	    // Condition to request disable send
	    #s_Ext_Req_Disable_Send := #i_External_Request.Request_Disable_Send;

	    // Condition to request disable receive
	    #s_Ext_Req_Disable_Recv := #i_External_Request.Request_Disable_Receive OR #i_Command.Man_Mode;

	    // Condition to request reset engergy saving
	    #s_Ext_Req_Rest_ESave := #i_External_Request.Request_Reset_EnergySave OR #io_Global.Common_Setting.Disable_Energy_Saving OR #i_Command.Cmd_Reset_ESave OR #s_FB_EQP_PEC_Position.s_PEC_Filter;

	    // Condition to request clear flow interface data
	    #s_Ext_Req_Clear_Data := #i_External_Request.Request_Clear_Data OR (#i_Command.Man_Clear AND #i_Command.Man_Mode);
	END_REGION

	REGION NETWORK DA: Equipment Layer - Basic
	    #s_FB_EQP_Transport(i_Enable                 := #io_System_Control.Enable,
	                        i_IO_Available           := #io_System_Control.IO_Available,
	                        i_Safety_OK              := #io_System_Control.Safety_OK,
	                        i_CMD_Reset              := #io_System_Control.OS_Reset,
	                        i_CMD_Start              := #io_System_Control.OS_Start,
	                        i_CMD_Controlled_Stop    := #io_System_Control.Controlled_Stop,
	                        i_End_PEC_Latch          := #s_PE_Position_Latch,
	                        i_Manual_Run             := #i_Command.Man_Run AND #i_Command.Man_Mode,
	                        i_CFG_Slave_Conveyor     := #i_Setting.Base_Conveyor.Slave_Mode,
	                        i_CFG_Enable_DieForward  := #i_Setting.Base_Conveyor.Enable_DieForward,
	                        i_Delay_Waiting_Item     := #i_Setting.Base_Conveyor.Delay_Waiting_Item,
	                        i_Delay_Dieback          := #i_Setting.Base_Conveyor.Delay_Dieback,
	                        i_Delay_Startup          := #i_Setting.Base_Conveyor.Delay_Startup,
	                        i_Delay_Finish_Handover  := #i_Setting.Base_Conveyor.Delay_Finish_Handover,
	                        i_Delay_Energysave       := #i_Setting.Base_Conveyor.Delay_Energysave,
	                        i_Delay_Cascade_Startup  := #i_Setting.Base_Conveyor.Delay_Cascade_Startup,
	                        i_Delay_Cascade_Shutdown := #i_Setting.Base_Conveyor.Delay_Cascade_Shutdown,
	                        i_Delay_Motor_Startup    := 0,
	                        i_Minimum_Gap            := #i_Setting.Flow_Control.Minimum_Gap,
	                        i_Minimum_Head_To_Head   := #i_Setting.Flow_Control.Minimum_Head_To_Head,
	                        i_Ext_Req_Stop           := #s_Ext_Req_Stop,
	                        i_Ext_Req_Halt           := #s_Ext_Req_Halt,
	                        i_Ext_Req_Dis_Send       := #s_Ext_Req_Disable_Send,
	                        i_Ext_Req_Dis_Recv       := #s_Ext_Req_Disable_Recv,
	                        i_Ext_Req_Rst_ESave      := #s_Ext_Req_Rest_ESave,
	                        i_Ext_Req_Clear_Data     := #s_Ext_Req_Clear_Data,
	                        o_Ready_To_Start         => #io_System_Control.Ready_To_Start,
	                        o_ST_Safety_Stop         => #o_General_Status.Safety_Stop,
	                        o_ST_Items               => #o_General_Status.Items,
	                        o_ST_Die_Back            => #o_General_Status.Die_Back,
	                        o_ST_Motor_Running       => #o_General_Status.Motor_Running,
	                        o_ST_Started             => #o_General_Status.Started,
	                        o_ST_Energy_Saving       => #o_General_Status.Energy_Saving,
	                        o_MTR_Run                => #s_CMD_Motor,
	                        io_Global                := #io_Global,
	                        io_FIF_Upstream          := #io_FIF_Upstream,
	                        io_FIF                   := #io_FIF,
	                        io_FIF_Downstream        := #io_FIF_Downstream);
	END_REGION

	REGION NETWORK EA: Hardware Layer - Interroll MultiControl 1
	    #s_Speed_Select := #i_External_Request.Request_Speed;

	    #s_FB_HW_MultiControl_U01(i_IO_Available            := #io_System_Control.IO_Available,
	                              i_Safety_OK               := #io_System_Control.Safety_OK,
	                              i_CMD_Reset               := #io_System_Control.OS_Reset,
	                              i_CMD_Clear_Stat          := #io_System_Control.OS_Clear_Statistics,
	                              i_HW_Setting              := #i_Setting.Hardware_U01,
	                              i_CFG_Motor_Switch_Time   := 500,
	                              i_CMD_Select_Speed        := #s_Speed_Select,
	                              i_CMD_Motor_Run           := #s_CMD_Motor,
	                              i_CMD_Motor_Reverse       := #s_CMD_Motor_Reverse,
	                              o_Ready_To_Reset          => #t_HW_VFD_U01_Ready_To_Reset,
	                              o_Req_Halt                => #s_HW_U01_Req_Halt,
	                              o_ER_Motor_1_Fault        => #t_ER_Motor_U01_Fault,
	                              o_ER_Motor_2_Fault        => #t_ER_Motor_U02_Fault,
	                              o_ER_Motor_3_Fault        => #t_ER_Motor_U03_Fault,
	                              o_ER_Motor_4_Fault        => #t_ER_Motor_U04_Fault,
	                              o_Speed_Selected          => #io_FIF.Speed,
	                              o_Diagnostics             => #o_Diagnostics.Hardware_U01,
	                              io_Global                 := #io_Global,
	                              io_MultiControl_Interface := #io_MultiControl_U01_IO);

	    IF #i_Setting.Hardware_U01.RD1_Motor_Number > 0 AND #i_Setting.Hardware_U01.RD1_Motor_Number <= 16 THEN
	        #t_ER_Motor_Fault[#i_Setting.Hardware_U01.RD1_Motor_Number] := #t_ER_Motor_U01_Fault;
	    END_IF;

	    IF #i_Setting.Hardware_U01.RD2_Motor_Number > 0 AND #i_Setting.Hardware_U01.RD2_Motor_Number <= 16 THEN
	        #t_ER_Motor_Fault[#i_Setting.Hardware_U01.RD2_Motor_Number] := #t_ER_Motor_U02_Fault;
	    END_IF;

	    IF #i_Setting.Hardware_U01.RD3_Motor_Number > 0 AND #i_Setting.Hardware_U01.RD3_Motor_Number <= 16 THEN
	        #t_ER_Motor_Fault[#i_Setting.Hardware_U01.RD3_Motor_Number] := #t_ER_Motor_U03_Fault;
	    END_IF;

	    IF #i_Setting.Hardware_U01.RD4_Motor_Number > 0 AND #i_Setting.Hardware_U01.RD4_Motor_Number <= 16 THEN
	        #t_ER_Motor_Fault[#i_Setting.Hardware_U01.RD4_Motor_Number] := #t_ER_Motor_U04_Fault;
	    END_IF;
	END_REGION

	REGION NETWORK EB: Hardware Layer - Interroll MultiControl 2
	    #s_Speed_Select := #i_External_Request.Request_Speed;

	    #s_FB_HW_MultiControl_U02(i_IO_Available            := #io_System_Control.IO_Available,
	                              i_Safety_OK               := #io_System_Control.Safety_OK,
	                              i_CMD_Reset               := #io_System_Control.OS_Reset,
	                              i_CMD_Clear_Stat          := #io_System_Control.OS_Clear_Statistics,
	                              i_HW_Setting              := #i_Setting.Hardware_U02,
	                              i_CFG_Motor_Switch_Time   := 500,
	                              i_CMD_Select_Speed        := #s_Speed_Select,
	                              i_CMD_Motor_Run           := #s_CMD_Motor,
	                              i_CMD_Motor_Reverse       := #s_CMD_Motor_Reverse,
	                              o_Ready_To_Reset          => #t_HW_VFD_U02_Ready_To_Reset,
	                              o_Req_Halt                => #s_HW_U02_Req_Halt,
	                              o_ER_Motor_1_Fault        => #t_ER_Motor_U01_Fault,
	                              o_ER_Motor_2_Fault        => #t_ER_Motor_U02_Fault,
	                              o_ER_Motor_3_Fault        => #t_ER_Motor_U03_Fault,
	                              o_ER_Motor_4_Fault        => #t_ER_Motor_U04_Fault,
	                              o_Diagnostics             => #o_Diagnostics.Hardware_U02,
	                              io_Global                 := #io_Global,
	                              io_MultiControl_Interface := #io_MultiControl_U02_IO);

	    IF #i_Setting.Hardware_U02.RD1_Motor_Number > 0 AND #i_Setting.Hardware_U02.RD1_Motor_Number <= 16 THEN
	        #t_ER_Motor_Fault[#i_Setting.Hardware_U02.RD1_Motor_Number] := #t_ER_Motor_U01_Fault;
	    END_IF;

	    IF #i_Setting.Hardware_U02.RD2_Motor_Number > 0 AND #i_Setting.Hardware_U02.RD2_Motor_Number <= 16 THEN
	        #t_ER_Motor_Fault[#i_Setting.Hardware_U02.RD2_Motor_Number] := #t_ER_Motor_U02_Fault;
	    END_IF;

	    IF #i_Setting.Hardware_U02.RD3_Motor_Number > 0 AND #i_Setting.Hardware_U02.RD3_Motor_Number <= 16 THEN
	        #t_ER_Motor_Fault[#i_Setting.Hardware_U02.RD3_Motor_Number] := #t_ER_Motor_U03_Fault;
	    END_IF;

	    IF #i_Setting.Hardware_U02.RD4_Motor_Number > 0 AND #i_Setting.Hardware_U02.RD4_Motor_Number <= 16 THEN
	        #t_ER_Motor_Fault[#i_Setting.Hardware_U02.RD4_Motor_Number] := #t_ER_Motor_U04_Fault;
	    END_IF;
	END_REGION

	REGION NETWORK EA: Hardware Layer - Interroll MultiControl 3
	    #s_Speed_Select := #i_External_Request.Request_Speed;

	    #s_FB_HW_MultiControl_U03(i_IO_Available            := #io_System_Control.IO_Available,
	                              i_Safety_OK               := #io_System_Control.Safety_OK,
	                              i_CMD_Reset               := #io_System_Control.OS_Reset,
	                              i_CMD_Clear_Stat          := #io_System_Control.OS_Clear_Statistics,
	                              i_HW_Setting              := #i_Setting.Hardware_U03,
	                              i_CFG_Motor_Switch_Time   := 500,
	                              i_CMD_Select_Speed        := #s_Speed_Select,
	                              i_CMD_Motor_Run           := #s_CMD_Motor,
	                              i_CMD_Motor_Reverse       := #s_CMD_Motor_Reverse,
	                              o_Ready_To_Reset          => #t_HW_VFD_U03_Ready_To_Reset,
	                              o_Req_Halt                => #s_HW_U03_Req_Halt,
	                              o_ER_Motor_1_Fault        => #t_ER_Motor_U01_Fault,
	                              o_ER_Motor_2_Fault        => #t_ER_Motor_U02_Fault,
	                              o_ER_Motor_3_Fault        => #t_ER_Motor_U03_Fault,
	                              o_ER_Motor_4_Fault        => #t_ER_Motor_U04_Fault,
	                              o_Diagnostics             => #o_Diagnostics.Hardware_U03,
	                              io_Global                 := #io_Global,
	                              io_MultiControl_Interface := #io_MultiControl_U03_IO);

	    IF #i_Setting.Hardware_U03.RD1_Motor_Number > 0 AND #i_Setting.Hardware_U03.RD1_Motor_Number <= 16 THEN
	        #t_ER_Motor_Fault[#i_Setting.Hardware_U03.RD1_Motor_Number] := #t_ER_Motor_U01_Fault;
	    END_IF;

	    IF #i_Setting.Hardware_U03.RD2_Motor_Number > 0 AND #i_Setting.Hardware_U03.RD2_Motor_Number <= 16 THEN
	        #t_ER_Motor_Fault[#i_Setting.Hardware_U03.RD2_Motor_Number] := #t_ER_Motor_U02_Fault;
	    END_IF;

	    IF #i_Setting.Hardware_U03.RD3_Motor_Number > 0 AND #i_Setting.Hardware_U03.RD3_Motor_Number <= 16 THEN
	        #t_ER_Motor_Fault[#i_Setting.Hardware_U03.RD3_Motor_Number] := #t_ER_Motor_U03_Fault;
	    END_IF;

	    IF #i_Setting.Hardware_U03.RD4_Motor_Number > 0 AND #i_Setting.Hardware_U03.RD4_Motor_Number <= 16 THEN
	        #t_ER_Motor_Fault[#i_Setting.Hardware_U03.RD4_Motor_Number] := #t_ER_Motor_U04_Fault;
	    END_IF;
	END_REGION

	REGION NETWORK EA: Hardware Layer - Interroll MultiControl 4
	    #s_Speed_Select := #i_External_Request.Request_Speed;

	    #s_FB_HW_MultiControl_U04(i_IO_Available            := #io_System_Control.IO_Available,
	                              i_Safety_OK               := #io_System_Control.Safety_OK,
	                              i_CMD_Reset               := #io_System_Control.OS_Reset,
	                              i_CMD_Clear_Stat          := #io_System_Control.OS_Clear_Statistics,
	                              i_HW_Setting              := #i_Setting.Hardware_U04,
	                              i_CFG_Motor_Switch_Time   := 500,
	                              i_CMD_Select_Speed        := #s_Speed_Select,
	                              i_CMD_Motor_Run           := #s_CMD_Motor,
	                              i_CMD_Motor_Reverse       := #s_CMD_Motor_Reverse,
	                              o_Ready_To_Reset          => #t_HW_VFD_U04_Ready_To_Reset,
	                              o_Req_Halt                => #s_HW_U04_Req_Halt,
	                              o_ER_Motor_1_Fault        => #t_ER_Motor_U01_Fault,
	                              o_ER_Motor_2_Fault        => #t_ER_Motor_U02_Fault,
	                              o_ER_Motor_3_Fault        => #t_ER_Motor_U03_Fault,
	                              o_ER_Motor_4_Fault        => #t_ER_Motor_U04_Fault,
	                              o_Diagnostics             => #o_Diagnostics.Hardware_U04,
	                              io_Global                 := #io_Global,
	                              io_MultiControl_Interface := #io_MultiControl_U04_IO);

	    IF #i_Setting.Hardware_U04.RD1_Motor_Number > 0 AND #i_Setting.Hardware_U04.RD1_Motor_Number <= 16 THEN
	        #t_ER_Motor_Fault[#i_Setting.Hardware_U04.RD1_Motor_Number] := #t_ER_Motor_U01_Fault;
	    END_IF;

	    IF #i_Setting.Hardware_U04.RD2_Motor_Number > 0 AND #i_Setting.Hardware_U04.RD2_Motor_Number <= 16 THEN
	        #t_ER_Motor_Fault[#i_Setting.Hardware_U04.RD2_Motor_Number] := #t_ER_Motor_U02_Fault;
	    END_IF;

	    IF #i_Setting.Hardware_U04.RD3_Motor_Number > 0 AND #i_Setting.Hardware_U04.RD3_Motor_Number <= 16 THEN
	        #t_ER_Motor_Fault[#i_Setting.Hardware_U04.RD3_Motor_Number] := #t_ER_Motor_U03_Fault;
	    END_IF;

	    IF #i_Setting.Hardware_U04.RD4_Motor_Number > 0 AND #i_Setting.Hardware_U04.RD4_Motor_Number <= 16 THEN
	        #t_ER_Motor_Fault[#i_Setting.Hardware_U04.RD4_Motor_Number] := #t_ER_Motor_U04_Fault;
	    END_IF;
	END_REGION

	REGION NETWORK: Copy Motor Alarm to Status

	    #o_Status.ER_Motor_1_Fault := #t_ER_Motor_Fault[1];
	    #o_Status.ER_Motor_2_Fault := #t_ER_Motor_Fault[2];
	    #o_Status.ER_Motor_3_Fault := #t_ER_Motor_Fault[3];
	    #o_Status.ER_Motor_4_Fault := #t_ER_Motor_Fault[4];
	    #o_Status.ER_Motor_5_Fault := #t_ER_Motor_Fault[5];
	    #o_Status.ER_Motor_6_Fault := #t_ER_Motor_Fault[6];
	    #o_Status.ER_Motor_7_Fault := #t_ER_Motor_Fault[7];
	    #o_Status.ER_Motor_8_Fault := #t_ER_Motor_Fault[8];
	    #o_Status.ER_Motor_9_Fault := #t_ER_Motor_Fault[9];
	    #o_Status.ER_Motor_10_Fault := #t_ER_Motor_Fault[10];
	    #o_Status.ER_Motor_11_Fault := #t_ER_Motor_Fault[11];
	    #o_Status.ER_Motor_12_Fault := #t_ER_Motor_Fault[12];
	    #o_Status.ER_Motor_13_Fault := #t_ER_Motor_Fault[13];
	    #o_Status.ER_Motor_14_Fault := #t_ER_Motor_Fault[14];
	    #o_Status.ER_Motor_15_Fault := #t_ER_Motor_Fault[15];
	    #o_Status.ER_Motor_16_Fault := #t_ER_Motor_Fault[16];

	END_REGION

	REGION NETWORK: Diagnositcs
	    #o_Diagnostics.RTS := #io_FIF.RTS;
	    #o_Diagnostics.TIP := #io_FIF.TIP;
	    #o_Diagnostics.Downstream_RTR := #io_FIF_Downstream.RTR;
	    #o_Diagnostics.Displacement := #io_FIF.Displacement;
	    #o_Diagnostics.Items_Count := MAX_UDINT(IN1 := #t_PEC_Position_Items, IN2 := #t_PEC_Trigger_Items);
	END_REGION

	REGION NETWORK FA: Make Generate Status
	    #o_Status.OL_Maintenance_Mode := #i_Command.Man_Mode;

	    #o_General_Status.Safety_Stop := NOT #io_System_Control.Safety_OK;
	    #o_General_Status.Off_Line := #o_Status.OL_Maintenance_Mode;
	    #o_General_Status.Manual := FALSE;
	    #o_General_Status.Error := #o_Status.ER_Motor_1_Fault
	    OR #o_Status.ER_Motor_2_Fault
	    OR #o_Status.ER_Motor_3_Fault
	    OR #o_Status.ER_Motor_4_Fault
	    OR #o_Status.ER_Motor_5_Fault
	    OR #o_Status.ER_Motor_6_Fault
	    OR #o_Status.ER_Motor_7_Fault
	    OR #o_Status.ER_Motor_8_Fault
	    OR #o_Status.ER_Motor_9_Fault
	    OR #o_Status.ER_Motor_10_Fault
	    OR #o_Status.ER_Motor_11_Fault
	    OR #o_Status.ER_Motor_12_Fault
	    OR #o_Status.ER_Motor_13_Fault
	    OR #o_Status.ER_Motor_14_Fault
	    OR #o_Status.ER_Motor_15_Fault
	    OR #o_Status.ER_Motor_16_Fault;
	    #o_General_Status.Jam := #o_Status.ER_PE1_Blockage OR #o_Status.ER_PE2_Blockage;
	END_REGION

	REGION NETWORK EA: System Feedback State
	    #io_System_Control.Ready_To_Reset := #t_PEC_Position_Ready_To_Reset
	    OR #t_PEC_Trigger_Ready_To_Reset
	    OR #t_HW_VFD_U01_Ready_To_Reset
	    OR #t_HW_VFD_U02_Ready_To_Reset
	    OR #t_HW_VFD_U03_Ready_To_Reset
	    OR #t_HW_VFD_U04_Ready_To_Reset;
	END_REGION
END_FUNCTION_BLOCK

TYPE "UDT_GL2S_IO"
VERSION : 0.1
   STRUCT
      IsCleared : Bool;
   END_STRUCT;

END_TYPE

TYPE "UDT_Conv_Triple_G115D_Status"
VERSION : 0.1
   STRUCT
      OL_Maintenance_Mode : Bool;   // Maintenance mode on
      ER_PE1_Blockage : Bool;   // PE1 blockage
      ER_PE2_Blockage : Bool;   // PE2 blockage
      ER_U01_VFD_PN_NotPresent : Bool;   // VFD 1# not present on profinet network
      ER_U01_VFD_PN_Error : Bool;   // VFD 1# has error profinet network
      ER_U01_VFD_Fault : Bool;   // VFD 1# has error
      WN_U01_VFD_Alarm : Bool;   // VFD 1# has an warning
      ER_U01_VFD_STO_Active : Bool;   // VFD 1# STO is active
      WN_U01_No_MemoryCard : Bool;   // Memory card is missing
      ER_U02_VFD_PN_NotPresent : Bool;   // VFD 2# not present on profinet network
      ER_U02_VFD_PN_Error : Bool;   // VFD 2# has error profinet network
      ER_U02_VFD_Fault : Bool;   // VFD 2# has error
      WN_U02_VFD_Alarm : Bool;   // VFD 2# has an warning
      ER_U02_VFD_STO_Active : Bool;   // VFD 2# STO is active
      WN_U02_No_MemoryCard : Bool;   // Memory card is missing
      ER_U03_VFD_PN_NotPresent : Bool;   // VFD 3# not present on profinet network
      ER_U03_VFD_PN_Error : Bool;   // VFD 3# has error profinet network
      ER_U03_VFD_Fault : Bool;   // VFD 3# has error
      WN_U03_VFD_Alarm : Bool;   // VFD 3# has an warning
      ER_U03_VFD_STO_Active : Bool;   // VFD 3# STO is active
      WN_U03_No_MemoryCard : Bool;   // Memory card is missing
      Spare_2_5 : Bool;   // Spare_2_5
      Spare_2_6 : Bool;   // Spare_2_6
      Spare_2_7 : Bool;   // Spare_2_7
      Spare_3_0 : Bool;   // Spare_3_0
      Spare_3_1 : Bool;   // Spare_3_1
      Spare_3_2 : Bool;   // Spare_3_2
      Spare_3_3 : Bool;   // Spare_3_3
      Spare_3_4 : Bool;   // Spare_3_4
      Spare_3_5 : Bool;   // Spare_3_5
      Spare_3_6 : Bool;   // Spare_3_6
      Spare_3_7 : Bool;   // Spare_3_7
      U01_FaultCode : Word;   // VFD 1# fault code
      U01_AlarmCode : Word;   // VFD 1# alarm code
      U02_FaultCode : Word;   // VFD 2# fault code
      U02_AlarmCode : Word;   // VFD 2# alarm code
      U03_FaultCode : Word;   // VFD 3# fault code
      U03_AlarmCode : Word;   // VFD 3# alarm code
   END_STRUCT;

END_TYPE

FUNCTION_BLOCK "FB_Conv_SWS"
{ S7_Optimized_Access := 'TRUE' }
VERSION : 0.1
   VAR_INPUT
      i_New_Item_Present : Bool;
      i_CMD_Divert_Left : Bool;
      i_CMD_Divert_Straight : Bool;
      i_CMD_Divert_Right : Bool;
      i_Setting : "UDT_Conv_SWS_Setting";
      i_External_Request : "UDT_External_Request";
      i_U401_Additional_HW_ID : HW_SUBMODULE;
      i_U401_Telegram_HW_ID : HW_SUBMODULE;
      i_U411_Additional_HW_ID : HW_SUBMODULE;
      i_U411_Telegram_HW_ID : HW_SUBMODULE;
      i_U421_Additional_HW_ID : HW_SUBMODULE;
      i_U421_Telegram_HW_ID : HW_SUBMODULE;
      i_U431_Additional_HW_ID : HW_SUBMODULE;
      i_U431_Telegram_HW_ID : HW_SUBMODULE;
      i_U441_Additional_HW_ID : HW_SUBMODULE;
      i_U441_Telegram_HW_ID : HW_SUBMODULE;
      i_U451_Additional_HW_ID : HW_SUBMODULE;
      i_U451_Telegram_HW_ID : HW_SUBMODULE;
      i_U461_Additional_HW_ID : HW_SUBMODULE;
      i_U461_Telegram_HW_ID : HW_SUBMODULE;
      i_U471_Additional_HW_ID : HW_SUBMODULE;
      i_U471_Telegram_HW_ID : HW_SUBMODULE;
      i_U481_Additional_HW_ID : HW_SUBMODULE;
      i_U481_Telegram_HW_ID : HW_SUBMODULE;
      i_Roller_Gateway_Input_HW_ID : HW_ANY;
      i_Roller_Gateway_Output_HW_ID : HW_ANY;
   END_VAR

   VAR_OUTPUT
      o_Status : "UDT_Conv_SWS_Status";
      o_General_Status : "UDT_General_Status";
   END_VAR

   VAR_IN_OUT
      io_Global : "UDT_Global";
      io_System_Control : "UDT_System_Control";
      io_Interface : "UDT_SWS_Interface";
      io_Gateway_Interface : "UDT_NT100_Interface";
      io_Command : "UDT_Conv_SWS_Command";
      io_FIF_Upstream : "UDT_Flow_Interface";
      io_FIF : "UDT_Flow_Interface";
      io_FIF_Downstream : "UDT_Flow_Interface";
   END_VAR

   VAR
      s_FB_Displacement_AccDec : "FB_Displacement_AccDec";
      s_FB_SWS_Roller_Interface : "FB_HW_SWS_Roller_Interface";
      s_FB_EQP_Transport : "FB_EQP_Transport";
      s_Trigger_FB_EQP_PEC_Position : "FB_EQP_PEC_Position";
      s_FB_SWS_Array_Control : "FB_SWS_Array_Control";
      s_U401_FB_SWS_EQP_Servo { S7_SetPoint := 'False'} : "FB_HW_SWS_S210";
      s_U411_FB_SWS_EQP_Servo { S7_SetPoint := 'False'} : "FB_HW_SWS_S210";
      s_U421_FB_SWS_EQP_Servo { S7_SetPoint := 'False'} : "FB_HW_SWS_S210";
      s_U431_FB_SWS_EQP_Servo { S7_SetPoint := 'False'} : "FB_HW_SWS_S210";
      s_U441_FB_SWS_EQP_Servo { S7_SetPoint := 'False'} : "FB_HW_SWS_S210";
      s_U451_FB_SWS_EQP_Servo { S7_SetPoint := 'False'} : "FB_HW_SWS_S210";
      s_U461_FB_SWS_EQP_Servo { S7_SetPoint := 'False'} : "FB_HW_SWS_S210";
      s_U471_FB_SWS_EQP_Servo { S7_SetPoint := 'False'} : "FB_HW_SWS_S210";
      s_U481_FB_SWS_EQP_Servo { S7_SetPoint := 'False'} : "FB_HW_SWS_S210";
      s_Servo_Array_Command : Array[1..#C_ARRAY_COUNT] of Struct
         CMD_Straight : Bool;
         CMD_Left : Bool;
         CMD_Right : Bool;
      END_STRUCT;
      s_Servo_Status { S7_SetPoint := 'False'} : Array[1..#C_ARRAY_COUNT] of "UDT_SWS_Servo_Status";
      s_Roller_Module_Status { ExternalAccessible := 'False'; ExternalVisible := 'False'; ExternalWritable := 'False'; S7_SetPoint := 'False'} : Array[1..9] of "UDT_SWS_Roller_Module_Status";
      s_Servo_Ready_To_Reset : Array[1..#C_ARRAY_COUNT] of Bool;
   END_VAR
   VAR RETAIN
      s_SW_Actual_Speed { S7_SetPoint := 'True'} : Int;
      s_CMD_Roller_Run : Bool;
      s_Ext_Req_Stop : Bool;
      s_Ext_Req_Halt : Bool;
      s_Ext_Req_Disable_Send : Bool;
      s_Ext_Req_Disable_Recv : Bool;
      s_Ext_Req_Rest_ESave : Bool;
      s_Ext_Req_Clear_Data : Bool;
   END_VAR

   VAR_TEMP
      t_GeoAddr {InstructionName := 'GEOADDR'; LibVersion := '1.0'} : GEOADDR;
      t_Ret_Val_Int : Int;   // Temp: Return Value Int
      t_Delayed_Item_Trigger : Bool;
   END_VAR

   VAR CONSTANT
      C_ARRAY_COUNT : UInt := 9;
   END_VAR


BEGIN
	REGION Conveyor Cycle Displacement
	    #io_FIF.Speed := #i_Setting.Hardware.Roller.Speed_Straight;

	    #s_FB_Displacement_AccDec(i_Conveyor_Speed   := #io_FIF.Speed,
	                              i_Accelaration     := #i_Setting.Hardware.Roller.Acceleration,
	                              i_Decelaration     := #i_Setting.Hardware.Roller.Deceleration,
	                              i_Prev_Cycle_Time  := #io_Global.OB_Prev_Cycle_Time,
	                              i_PPI_Displacement := 0,
	                              i_Section_Run      := #io_FIF.Motor_Run,
	                              o_Motor_On_Speed   => #o_General_Status.Motor_On_Speed,
	                              o_Motor_Stopped    => #io_FIF.Motor_Stopped,
	                              o_Actual_Speed     => #s_SW_Actual_Speed,
	                              o_Displacement     => #io_FIF.Displacement);

	    #o_General_Status.Motor_Stopped := #io_FIF.Motor_Stopped;
	END_REGION

	REGION Roller Hardware Interface
	    #s_FB_SWS_Roller_Interface(i_CFG_HW_Port                := #i_Roller_Gateway_Input_HW_ID,
	                               i_IO_Available               := #io_System_Control.IO_Available,
	                               i_OB_First_Scan              := #io_Global.OS_First_Scan,
	                               i_CMD_Reset                  := #io_System_Control.OS_Reset,
	                               i_CFG_Status_Interval        := #i_Setting.Roller_Interface.Status_Interval,
	                               i_CFG_Num_Of_Comm_Error      := #i_Setting.Roller_Interface.Num_Of_Comm_Error,
	                               i_Sett_Roller_Hardware       := #i_Setting.Hardware.Roller,
	                               i_Roller_Running             := #io_FIF.Motor_Run,
	                               o_ER_Modbus_Initialize_Fault => #o_Status.ER_Modbus_Gateway_Initialize_Fault,
	                               o_ER_Modbus_Com_Error        => #o_Status.ER_Modbus_Gateway_Communication_Fault,
	                               o_Modules_Status             => #s_Roller_Module_Status);

	END_REGION

	REGION Conditions to basic control
	    // Condition to request stop
	    #s_Ext_Req_Stop := #s_Servo_Status[1].ER_PN_NotPresent
	    OR #s_Servo_Status[2].ER_PN_NotPresent
	    OR #s_Servo_Status[3].ER_PN_NotPresent
	    OR #s_Servo_Status[4].ER_PN_NotPresent
	    OR #s_Servo_Status[5].ER_PN_NotPresent
	    OR #s_Servo_Status[6].ER_PN_NotPresent
	    OR #s_Servo_Status[7].ER_PN_NotPresent
	    OR #s_Servo_Status[8].ER_PN_NotPresent
	    OR #s_Servo_Status[9].ER_PN_NotPresent
	    OR #s_Servo_Status[1].ER_Servo_Fault
	    OR #s_Servo_Status[2].ER_Servo_Fault
	    OR #s_Servo_Status[3].ER_Servo_Fault
	    OR #s_Servo_Status[4].ER_Servo_Fault
	    OR #s_Servo_Status[5].ER_Servo_Fault
	    OR #s_Servo_Status[6].ER_Servo_Fault
	    OR #s_Servo_Status[7].ER_Servo_Fault
	    OR #s_Servo_Status[8].ER_Servo_Fault
	    OR #s_Servo_Status[9].ER_Servo_Fault
	    OR #s_Servo_Status[1].ER_Home_Position_Missed
	    OR #s_Servo_Status[2].ER_Home_Position_Missed
	    OR #s_Servo_Status[3].ER_Home_Position_Missed
	    OR #s_Servo_Status[4].ER_Home_Position_Missed
	    OR #s_Servo_Status[5].ER_Home_Position_Missed
	    OR #s_Servo_Status[6].ER_Home_Position_Missed
	    OR #s_Servo_Status[7].ER_Home_Position_Missed
	    OR #s_Servo_Status[8].ER_Home_Position_Missed
	    OR #s_Servo_Status[9].ER_Home_Position_Missed
	    OR #s_Servo_Status[1].ER_STO_Active
	    OR #s_Servo_Status[2].ER_STO_Active
	    OR #s_Servo_Status[3].ER_STO_Active
	    OR #s_Servo_Status[4].ER_STO_Active
	    OR #s_Servo_Status[5].ER_STO_Active
	    OR #s_Servo_Status[6].ER_STO_Active
	    OR #s_Servo_Status[7].ER_STO_Active
	    OR #s_Servo_Status[8].ER_STO_Active
	    OR #s_Servo_Status[9].ER_STO_Active
	    OR #i_External_Request.Request_Stop;

	    // Condition to request halt
	    #s_Ext_Req_Halt := #i_External_Request.Request_Halt OR #io_Command.Man_Mode;

	    // Condition to request disable send
	    #s_Ext_Req_Disable_Send := #i_External_Request.Request_Disable_Send;

	    // Condition to request disable receive
	    #s_Ext_Req_Disable_Recv := #i_External_Request.Request_Disable_Receive OR #io_Command.Man_Mode;

	    // Condition to request reset engergy saving
	    #s_Ext_Req_Rest_ESave := #i_External_Request.Request_Reset_EnergySave OR #io_Global.Common_Setting.Disable_Energy_Saving OR #io_Command.Cmd_Reset_ESave;

	    // Condition to request clear flow interface data
	    #s_Ext_Req_Clear_Data := #i_External_Request.Request_Clear_Data OR (#io_Command.Man_Clear AND #io_Command.Man_Mode);
	END_REGION

	REGION Roller Equipment Control

	    #s_FB_EQP_Transport(i_Enable                := #io_System_Control.Enable,
	                        i_IO_Available          := #io_System_Control.IO_Available,
	                        i_Safety_OK             := #io_System_Control.Safety_OK,
	                        i_CMD_Reset             := #io_System_Control.OS_Reset,
	                        i_CMD_Start             := #io_System_Control.OS_Start,
	                        i_CMD_Controlled_Stop   := #io_System_Control.Controlled_Stop,
	                        i_End_PEC_Latch         := FALSE,
	                        i_Manual_Run            := #io_Command.Man_Run AND #io_Command.Man_Mode,
	                        i_CFG_Slave_Conveyor    := #i_Setting.Base_Conveyor.Slave_Mode,
	                        i_CFG_Enable_DieForward := #i_Setting.Base_Conveyor.Enable_DieForward,
	                        i_Delay_Waiting_Item    := #i_Setting.Base_Conveyor.Delay_Waiting_Item,
	                        i_Delay_Dieback         := #i_Setting.Base_Conveyor.Delay_Dieback,
	                        i_Delay_Finish_Handover := #i_Setting.Base_Conveyor.Delay_Finish_Handover,
	                        i_Delay_Energysave      := #i_Setting.Base_Conveyor.Delay_Energysave,
	                        i_Delay_Cascade_Startup := #i_Setting.Base_Conveyor.Delay_Cascade_Startup,
	                        i_Delay_Startup         := #i_Setting.Base_Conveyor.Delay_Startup,
	                        i_Delay_Motor_Startup   := 0,
	                        i_Minimum_Gap           := 0,
	                        i_Minimum_Head_To_Head  := 0,
	                        i_Ext_Req_Stop          := #s_Ext_Req_Stop,
	                        i_Ext_Req_Halt          := #s_Ext_Req_Halt,
	                        i_Ext_Req_Dis_Send      := #s_Ext_Req_Disable_Send,
	                        i_Ext_Req_Dis_Recv      := #s_Ext_Req_Disable_Recv,
	                        i_Ext_Req_Rst_ESave     := #s_Ext_Req_Rest_ESave,
	                        i_Ext_Req_Clear_Data    := #s_Ext_Req_Clear_Data,
	                        o_Ready_To_Start        => #io_System_Control.Ready_To_Start,
	                        o_ST_Safety_Stop        => #o_General_Status.Safety_Stop,
	                        o_ST_Items              => #o_General_Status.Items,
	                        o_ST_Die_Back           => #o_General_Status.Die_Back,
	                        o_ST_Motor_Running      => #o_General_Status.Motor_Running,
	                        o_ST_Started            => #o_General_Status.Started,
	                        o_ST_Energy_Saving      => #o_General_Status.Energy_Saving,
	                        o_MTR_Run               => #s_CMD_Roller_Run,
	                        io_Global               := #io_Global,
	                        io_FIF_Upstream         := #io_FIF_Upstream,
	                        io_FIF                  := #io_FIF,
	                        io_FIF_Downstream       := #io_FIF_Downstream);

	END_REGION

	REGION Servo Array Control

	    #s_FB_SWS_Array_Control(i_CMD_Roller_Run       := #s_CMD_Roller_Run,
	                            i_CMD_Straight         := NOT #i_CMD_Divert_Left AND NOT #i_CMD_Divert_Right,
	                            i_CMD_Divert_Left      := #i_CMD_Divert_Left,
	                            i_CMD_Divert_Right     := #i_CMD_Divert_Right,
	                            i_CMD_Manual_Mode      := #io_Command.Manual_Mode,
	                            i_CMD_Fixed_Straight   := #io_Command.Manual_Fixed_Straight,
	                            i_CMD_Fixed_Left       := #io_Command.Manual_Fixed_Left,
	                            i_CMD_Fixed_Right      := #io_Command.Manual_Fixed_Right,
	                            i_CMD_Fixed_Ratio      := #io_Command.Manual_Fixed_Ratio,
	                            i_New_Item_Present     := #t_Delayed_Item_Trigger,
	                            i_Cycle_Count          := #io_FIF.Displacement,
	                            i_Setting              := #i_Setting.Divert,
	                            i_Servos_Status        := #s_Servo_Status,
	                            io_Global              := #io_Global,
	                            io_Array_Command       := #s_Servo_Array_Command,
	                            io_Roller_IO_Interface := #io_Interface.Roller_Module);
	END_REGION

	REGION Servo Switch Hardware Interface
	    REGION U401 Servo
	        #s_U401_FB_SWS_EQP_Servo(i_Additional_HW_ID         := #i_U401_Additional_HW_ID,
	                                 i_Telegram_HW_ID           := #i_U401_Telegram_HW_ID,
	                                 i_IO_Available             := #io_System_Control.IO_Available,
	                                 i_Safety_OK                := #io_System_Control.Safety_OK,
	                                 i_CMD_Reset                := #io_System_Control.OS_Reset,
	                                 i_CMD_Maintenance_Mode     := #io_Command.Man_Mode_Servo,
	                                 i_CMD_Disable_Axis         := #io_Command.Servo_Array[1].Man_Disable_Axis,
	                                 i_CMD_Home                 := #io_Command.Servo_Array[1].Man_Home,
	                                 i_CMD_Jog_Left             := #io_Command.Servo_Array[1].Man_Jog_Left,
	                                 i_CMD_Jog_Right            := #io_Command.Servo_Array[1].Man_Jog_Right,
	                                 i_CMD_Save                 := #io_Command.Servo_Array[1].Man_Save_Parameter,
	                                 i_CMD_Straight             := #s_Servo_Array_Command[1].CMD_Straight,
	                                 i_CMD_Divert_Left          := #s_Servo_Array_Command[1].CMD_Left,
	                                 i_CMD_Divert_Right         := #s_Servo_Array_Command[1].CMD_Right,
	                                 i_HW_Setting               := #i_Setting.Hardware.Servo_U401,
	                                 o_Ready_To_Reset           => #s_Servo_Ready_To_Reset[1],
	                                 o_ER_PN_Not_Present        => #s_Servo_Status[1].ER_PN_NotPresent,
	                                 o_ER_PN_Error              => #s_Servo_Status[1].ER_PN_Error,
	                                 o_ST_Axis_Enabled          => #s_Servo_Status[1].ST_Axis_Enabled,
	                                 o_ST_Position_Reached      => #s_Servo_Status[1].ST_Axis_Position_Reached,
	                                 o_OL_Maintenance_Mode      => #s_Servo_Status[1].OL_Maintenance_Mode,
	                                 o_ER_STO_Active            => #s_Servo_Status[1].ER_STO_Active,
	                                 o_WN_Motor_Alarm           => #s_Servo_Status[1].WN_Servo_Warn,
	                                 o_ER_Motor_Fault           => #s_Servo_Status[1].ER_Servo_Fault,
	                                 o_ER_Home_Position_Missing => #s_Servo_Status[1].ER_Home_Position_Missed,
	                                 o_ST_Act_Position          => #s_Servo_Status[1].ST_Act_Position,
	                                 o_AlarmCode                 => #s_Servo_Status[1].AlarmCode,
	                                 o_FaultCode                => #s_Servo_Status[1].ErrorCode,
	                                 io_Global                  := #io_Global,
	                                 io_S210_Interface          := #io_Interface.Servo1);
	    END_REGION

	    REGION U411 Servo
	        #s_U411_FB_SWS_EQP_Servo(i_Telegram_HW_ID           := #i_U411_Telegram_HW_ID,
	                                 i_Additional_HW_ID         := #i_U411_Additional_HW_ID,
	                                 i_IO_Available             := #io_System_Control.IO_Available,
	                                 i_Safety_OK                := #io_System_Control.Safety_OK,
	                                 i_CMD_Reset                := #io_System_Control.OS_Reset,
	                                 i_CMD_Maintenance_Mode     := #io_Command.Man_Mode_Servo,
	                                 i_CMD_Disable_Axis         := #io_Command.Servo_Array[2].Man_Disable_Axis,
	                                 i_CMD_Home                 := #io_Command.Servo_Array[2].Man_Home,
	                                 i_CMD_Jog_Left             := #io_Command.Servo_Array[2].Man_Jog_Left,
	                                 i_CMD_Jog_Right            := #io_Command.Servo_Array[2].Man_Jog_Right,
	                                 i_CMD_Save                 := #io_Command.Servo_Array[2].Man_Save_Parameter,
	                                 i_CMD_Straight             := #s_Servo_Array_Command[2].CMD_Straight,
	                                 i_CMD_Divert_Left          := #s_Servo_Array_Command[2].CMD_Left,
	                                 i_CMD_Divert_Right         := #s_Servo_Array_Command[2].CMD_Right,
	                                 i_HW_Setting               := #i_Setting.Hardware.Servo_U411,
	                                 o_Ready_To_Reset           => #s_Servo_Ready_To_Reset[2],
	                                 o_ER_PN_Not_Present        => #s_Servo_Status[2].ER_PN_NotPresent,
	                                 o_ER_PN_Error              => #s_Servo_Status[2].ER_PN_Error,
	                                 o_ST_Axis_Enabled          => #s_Servo_Status[2].ST_Axis_Enabled,
	                                 o_ST_Position_Reached      => #s_Servo_Status[2].ST_Axis_Position_Reached,
	                                 o_OL_Maintenance_Mode      => #s_Servo_Status[2].OL_Maintenance_Mode,
	                                 o_ER_STO_Active            => #s_Servo_Status[2].ER_STO_Active,
	                                 o_WN_Motor_Alarm           => #s_Servo_Status[2].WN_Servo_Warn,
	                                 o_ER_Motor_Fault           => #s_Servo_Status[2].ER_Servo_Fault,
	                                 o_ER_Home_Position_Missing => #s_Servo_Status[2].ER_Home_Position_Missed,
	                                 o_ST_Act_Position          => #s_Servo_Status[2].ST_Act_Position,
	                                 o_AlarmCode                 => #s_Servo_Status[2].AlarmCode,
	                                 o_FaultCode                => #s_Servo_Status[2].ErrorCode,
	                                 io_Global                  := #io_Global,
	                                 io_S210_Interface          := #io_Interface.Servo2);
	    END_REGION

	    REGION U421 Servo
	        #s_U421_FB_SWS_EQP_Servo(i_Telegram_HW_ID           := #i_U421_Telegram_HW_ID,
	                                 i_Additional_HW_ID         := #i_U421_Additional_HW_ID,
	                                 i_IO_Available             := #io_System_Control.IO_Available,
	                                 i_Safety_OK                := #io_System_Control.Safety_OK,
	                                 i_CMD_Reset                := #io_System_Control.OS_Reset,
	                                 i_CMD_Maintenance_Mode     := #io_Command.Man_Mode_Servo,
	                                 i_CMD_Disable_Axis         := #io_Command.Servo_Array[3].Man_Disable_Axis,
	                                 i_CMD_Home                 := #io_Command.Servo_Array[3].Man_Home,
	                                 i_CMD_Jog_Left             := #io_Command.Servo_Array[3].Man_Jog_Left,
	                                 i_CMD_Jog_Right            := #io_Command.Servo_Array[3].Man_Jog_Right,
	                                 i_CMD_Save                 := #io_Command.Servo_Array[3].Man_Save_Parameter,
	                                 i_CMD_Straight             := #s_Servo_Array_Command[3].CMD_Straight,
	                                 i_CMD_Divert_Left          := #s_Servo_Array_Command[3].CMD_Left,
	                                 i_CMD_Divert_Right         := #s_Servo_Array_Command[3].CMD_Right,
	                                 i_HW_Setting               := #i_Setting.Hardware.Servo_U421,
	                                 o_Ready_To_Reset           => #s_Servo_Ready_To_Reset[3],
	                                 o_ER_PN_Not_Present        => #s_Servo_Status[3].ER_PN_NotPresent,
	                                 o_ER_PN_Error              => #s_Servo_Status[3].ER_PN_Error,
	                                 o_ST_Axis_Enabled          => #s_Servo_Status[3].ST_Axis_Enabled,
	                                 o_ST_Position_Reached      => #s_Servo_Status[3].ST_Axis_Position_Reached,
	                                 o_OL_Maintenance_Mode      => #s_Servo_Status[3].OL_Maintenance_Mode,
	                                 o_ER_STO_Active            => #s_Servo_Status[3].ER_STO_Active,
	                                 o_WN_Motor_Alarm           => #s_Servo_Status[3].WN_Servo_Warn,
	                                 o_ER_Motor_Fault           => #s_Servo_Status[3].ER_Servo_Fault,
	                                 o_ER_Home_Position_Missing => #s_Servo_Status[3].ER_Home_Position_Missed,
	                                 o_ST_Act_Position          => #s_Servo_Status[3].ST_Act_Position,
	                                 o_AlarmCode                 => #s_Servo_Status[3].AlarmCode,
	                                 o_FaultCode                => #s_Servo_Status[3].ErrorCode,
	                                 io_Global                  := #io_Global,
	                                 io_S210_Interface          := #io_Interface.Servo3);
	    END_REGION

	    REGION U431 Servo
	        #s_U431_FB_SWS_EQP_Servo(i_Telegram_HW_ID           := #i_U431_Telegram_HW_ID,
	                                 i_Additional_HW_ID         := #i_U431_Additional_HW_ID,
	                                 i_IO_Available             := #io_System_Control.IO_Available,
	                                 i_Safety_OK                := #io_System_Control.Safety_OK,
	                                 i_CMD_Reset                := #io_System_Control.OS_Reset,
	                                 i_CMD_Maintenance_Mode     := #io_Command.Man_Mode_Servo,
	                                 i_CMD_Disable_Axis         := #io_Command.Servo_Array[4].Man_Disable_Axis,
	                                 i_CMD_Home                 := #io_Command.Servo_Array[4].Man_Home,
	                                 i_CMD_Jog_Left             := #io_Command.Servo_Array[4].Man_Jog_Left,
	                                 i_CMD_Jog_Right            := #io_Command.Servo_Array[4].Man_Jog_Right,
	                                 i_CMD_Save                 := #io_Command.Servo_Array[5].Man_Save_Parameter,
	                                 i_CMD_Straight             := #s_Servo_Array_Command[4].CMD_Straight,
	                                 i_CMD_Divert_Left          := #s_Servo_Array_Command[4].CMD_Left,
	                                 i_CMD_Divert_Right         := #s_Servo_Array_Command[4].CMD_Right,
	                                 i_HW_Setting               := #i_Setting.Hardware.Servo_U431,
	                                 o_Ready_To_Reset           => #s_Servo_Ready_To_Reset[4],
	                                 o_ER_PN_Not_Present        => #s_Servo_Status[4].ER_PN_NotPresent,
	                                 o_ER_PN_Error              => #s_Servo_Status[4].ER_PN_Error,
	                                 o_ST_Axis_Enabled          => #s_Servo_Status[4].ST_Axis_Enabled,
	                                 o_ST_Position_Reached      => #s_Servo_Status[4].ST_Axis_Position_Reached,
	                                 o_OL_Maintenance_Mode      => #s_Servo_Status[4].OL_Maintenance_Mode,
	                                 o_ER_STO_Active            => #s_Servo_Status[4].ER_STO_Active,
	                                 o_WN_Motor_Alarm           => #s_Servo_Status[4].WN_Servo_Warn,
	                                 o_ER_Motor_Fault           => #s_Servo_Status[4].ER_Servo_Fault,
	                                 o_ER_Home_Position_Missing => #s_Servo_Status[4].ER_Home_Position_Missed,
	                                 o_ST_Act_Position          => #s_Servo_Status[4].ST_Act_Position,
	                                 o_AlarmCode                 => #s_Servo_Status[4].AlarmCode,
	                                 o_FaultCode                => #s_Servo_Status[4].ErrorCode,
	                                 io_Global                  := #io_Global,
	                                 io_S210_Interface          := #io_Interface.Servo4);
	    END_REGION

	    REGION U441 Servo
	        #s_U441_FB_SWS_EQP_Servo(i_Telegram_HW_ID           := #i_U441_Telegram_HW_ID,
	                                 i_Additional_HW_ID         := #i_U441_Additional_HW_ID,
	                                 i_IO_Available             := #io_System_Control.IO_Available,
	                                 i_Safety_OK                := #io_System_Control.Safety_OK,
	                                 i_CMD_Reset                := #io_System_Control.OS_Reset,
	                                 i_CMD_Maintenance_Mode     := #io_Command.Man_Mode_Servo,
	                                 i_CMD_Disable_Axis         := #io_Command.Servo_Array[5].Man_Disable_Axis,
	                                 i_CMD_Home                 := #io_Command.Servo_Array[5].Man_Home,
	                                 i_CMD_Jog_Left             := #io_Command.Servo_Array[5].Man_Jog_Left,
	                                 i_CMD_Jog_Right            := #io_Command.Servo_Array[5].Man_Jog_Right,
	                                 i_CMD_Save                 := #io_Command.Servo_Array[5].Man_Save_Parameter,
	                                 i_CMD_Straight             := #s_Servo_Array_Command[5].CMD_Straight,
	                                 i_CMD_Divert_Left          := #s_Servo_Array_Command[5].CMD_Left,
	                                 i_CMD_Divert_Right         := #s_Servo_Array_Command[5].CMD_Right,
	                                 i_HW_Setting               := #i_Setting.Hardware.Servo_U441,
	                                 o_Ready_To_Reset           => #s_Servo_Ready_To_Reset[5],
	                                 o_ER_PN_Not_Present        => #s_Servo_Status[5].ER_PN_NotPresent,
	                                 o_ER_PN_Error              => #s_Servo_Status[5].ER_PN_Error,
	                                 o_ST_Axis_Enabled          => #s_Servo_Status[5].ST_Axis_Enabled,
	                                 o_ST_Position_Reached      => #s_Servo_Status[5].ST_Axis_Position_Reached,
	                                 o_OL_Maintenance_Mode      => #s_Servo_Status[5].OL_Maintenance_Mode,
	                                 o_ER_STO_Active            => #s_Servo_Status[5].ER_STO_Active,
	                                 o_WN_Motor_Alarm           => #s_Servo_Status[5].WN_Servo_Warn,
	                                 o_ER_Motor_Fault           => #s_Servo_Status[5].ER_Servo_Fault,
	                                 o_ER_Home_Position_Missing => #s_Servo_Status[5].ER_Home_Position_Missed,
	                                 o_ST_Act_Position          => #s_Servo_Status[5].ST_Act_Position,
	                                 o_AlarmCode                 => #s_Servo_Status[5].AlarmCode,
	                                 o_FaultCode                => #s_Servo_Status[5].ErrorCode,
	                                 io_Global                  := #io_Global,
	                                 io_S210_Interface          := #io_Interface.Servo5);
	    END_REGION

	    REGION U451 Servo
	        #s_U451_FB_SWS_EQP_Servo(i_Telegram_HW_ID           := #i_U451_Telegram_HW_ID,
	                                 i_Additional_HW_ID         := #i_U451_Additional_HW_ID,
	                                 i_IO_Available             := #io_System_Control.IO_Available,
	                                 i_Safety_OK                := #io_System_Control.Safety_OK,
	                                 i_CMD_Reset                := #io_System_Control.OS_Reset,
	                                 i_CMD_Maintenance_Mode     := #io_Command.Man_Mode_Servo,
	                                 i_CMD_Disable_Axis         := #io_Command.Servo_Array[6].Man_Disable_Axis,
	                                 i_CMD_Home                 := #io_Command.Servo_Array[6].Man_Home,
	                                 i_CMD_Jog_Left             := #io_Command.Servo_Array[6].Man_Jog_Left,
	                                 i_CMD_Jog_Right            := #io_Command.Servo_Array[6].Man_Jog_Right,
	                                 i_CMD_Save                 := #io_Command.Servo_Array[6].Man_Save_Parameter,
	                                 i_CMD_Straight             := #s_Servo_Array_Command[6].CMD_Straight,
	                                 i_CMD_Divert_Left          := #s_Servo_Array_Command[6].CMD_Left,
	                                 i_CMD_Divert_Right         := #s_Servo_Array_Command[6].CMD_Right,
	                                 i_HW_Setting               := #i_Setting.Hardware.Servo_U451,
	                                 o_Ready_To_Reset           => #s_Servo_Ready_To_Reset[6],
	                                 o_ER_PN_Not_Present        => #s_Servo_Status[6].ER_PN_NotPresent,
	                                 o_ER_PN_Error              => #s_Servo_Status[6].ER_PN_Error,
	                                 o_ST_Axis_Enabled          => #s_Servo_Status[6].ST_Axis_Enabled,
	                                 o_ST_Position_Reached      => #s_Servo_Status[6].ST_Axis_Position_Reached,
	                                 o_OL_Maintenance_Mode      => #s_Servo_Status[6].OL_Maintenance_Mode,
	                                 o_ER_STO_Active            => #s_Servo_Status[6].ER_STO_Active,
	                                 o_WN_Motor_Alarm           => #s_Servo_Status[6].WN_Servo_Warn,
	                                 o_ER_Motor_Fault           => #s_Servo_Status[6].ER_Servo_Fault,
	                                 o_ER_Home_Position_Missing => #s_Servo_Status[6].ER_Home_Position_Missed,
	                                 o_ST_Act_Position          => #s_Servo_Status[6].ST_Act_Position,
	                                 o_AlarmCode                 => #s_Servo_Status[6].AlarmCode,
	                                 o_FaultCode                => #s_Servo_Status[6].ErrorCode,
	                                 io_Global                  := #io_Global,
	                                 io_S210_Interface          := #io_Interface.Servo6);
	    END_REGION

	    REGION U461 Servo
	        #s_U461_FB_SWS_EQP_Servo(i_Telegram_HW_ID           := #i_U461_Telegram_HW_ID,
	                                 i_Additional_HW_ID         := #i_U461_Additional_HW_ID,
	                                 i_IO_Available             := #io_System_Control.IO_Available,
	                                 i_Safety_OK                := #io_System_Control.Safety_OK,
	                                 i_CMD_Reset                := #io_System_Control.OS_Reset,
	                                 i_CMD_Maintenance_Mode     := #io_Command.Man_Mode_Servo,
	                                 i_CMD_Disable_Axis         := #io_Command.Servo_Array[7].Man_Disable_Axis,
	                                 i_CMD_Home                 := #io_Command.Servo_Array[7].Man_Home,
	                                 i_CMD_Jog_Left             := #io_Command.Servo_Array[7].Man_Jog_Left,
	                                 i_CMD_Jog_Right            := #io_Command.Servo_Array[7].Man_Jog_Right,
	                                 i_CMD_Save                 := #io_Command.Servo_Array[7].Man_Save_Parameter,
	                                 i_CMD_Straight             := #s_Servo_Array_Command[7].CMD_Straight,
	                                 i_CMD_Divert_Left          := #s_Servo_Array_Command[7].CMD_Left,
	                                 i_CMD_Divert_Right         := #s_Servo_Array_Command[7].CMD_Right,
	                                 i_HW_Setting               := #i_Setting.Hardware.Servo_U461,
	                                 o_Ready_To_Reset           => #s_Servo_Ready_To_Reset[7],
	                                 o_ER_PN_Not_Present        => #s_Servo_Status[7].ER_PN_NotPresent,
	                                 o_ER_PN_Error              => #s_Servo_Status[7].ER_PN_Error,
	                                 o_ST_Axis_Enabled          => #s_Servo_Status[7].ST_Axis_Enabled,
	                                 o_ST_Position_Reached      => #s_Servo_Status[7].ST_Axis_Position_Reached,
	                                 o_OL_Maintenance_Mode      => #s_Servo_Status[7].OL_Maintenance_Mode,
	                                 o_ER_STO_Active            => #s_Servo_Status[7].ER_STO_Active,
	                                 o_WN_Motor_Alarm           => #s_Servo_Status[7].WN_Servo_Warn,
	                                 o_ER_Motor_Fault           => #s_Servo_Status[7].ER_Servo_Fault,
	                                 o_ER_Home_Position_Missing => #s_Servo_Status[7].ER_Home_Position_Missed,
	                                 o_ST_Act_Position          => #s_Servo_Status[7].ST_Act_Position,
	                                 o_AlarmCode                 => #s_Servo_Status[7].AlarmCode,
	                                 o_FaultCode                => #s_Servo_Status[7].ErrorCode,
	                                 io_Global                  := #io_Global,
	                                 io_S210_Interface          := #io_Interface.Servo7);
	    END_REGION

	    REGION U471 Servo
	        #s_U471_FB_SWS_EQP_Servo(i_Telegram_HW_ID           := #i_U471_Telegram_HW_ID,
	                                 i_Additional_HW_ID         := #i_U471_Additional_HW_ID,
	                                 i_IO_Available             := #io_System_Control.IO_Available,
	                                 i_Safety_OK                := #io_System_Control.Safety_OK,
	                                 i_CMD_Reset                := #io_System_Control.OS_Reset,
	                                 i_CMD_Maintenance_Mode     := #io_Command.Man_Mode_Servo,
	                                 i_CMD_Disable_Axis         := #io_Command.Servo_Array[8].Man_Disable_Axis,
	                                 i_CMD_Home                 := #io_Command.Servo_Array[8].Man_Home,
	                                 i_CMD_Jog_Left             := #io_Command.Servo_Array[8].Man_Jog_Left,
	                                 i_CMD_Jog_Right            := #io_Command.Servo_Array[8].Man_Jog_Right,
	                                 i_CMD_Save                 := #io_Command.Servo_Array[8].Man_Save_Parameter,
	                                 i_CMD_Straight             := #s_Servo_Array_Command[8].CMD_Straight,
	                                 i_CMD_Divert_Left          := #s_Servo_Array_Command[8].CMD_Left,
	                                 i_CMD_Divert_Right         := #s_Servo_Array_Command[8].CMD_Right,
	                                 i_HW_Setting               := #i_Setting.Hardware.Servo_U471,
	                                 o_Ready_To_Reset           => #s_Servo_Ready_To_Reset[8],
	                                 o_ER_PN_Not_Present        => #s_Servo_Status[8].ER_PN_NotPresent,
	                                 o_ER_PN_Error              => #s_Servo_Status[8].ER_PN_Error,
	                                 o_ST_Axis_Enabled          => #s_Servo_Status[8].ST_Axis_Enabled,
	                                 o_ST_Position_Reached      => #s_Servo_Status[8].ST_Axis_Position_Reached,
	                                 o_OL_Maintenance_Mode      => #s_Servo_Status[8].OL_Maintenance_Mode,
	                                 o_ER_STO_Active            => #s_Servo_Status[8].ER_STO_Active,
	                                 o_WN_Motor_Alarm           => #s_Servo_Status[8].WN_Servo_Warn,
	                                 o_ER_Motor_Fault           => #s_Servo_Status[8].ER_Servo_Fault,
	                                 o_ER_Home_Position_Missing => #s_Servo_Status[8].ER_Home_Position_Missed,
	                                 o_ST_Act_Position          => #s_Servo_Status[8].ST_Act_Position,
	                                 o_AlarmCode                 => #s_Servo_Status[8].AlarmCode,
	                                 o_FaultCode                => #s_Servo_Status[8].ErrorCode,
	                                 io_Global                  := #io_Global,
	                                 io_S210_Interface          := #io_Interface.Servo8);
	    END_REGION

	    REGION U481 Servo
	        #s_U481_FB_SWS_EQP_Servo(i_Telegram_HW_ID           := #i_U481_Telegram_HW_ID,
	                                 i_Additional_HW_ID         := #i_U481_Additional_HW_ID,
	                                 i_IO_Available             := #io_System_Control.IO_Available,
	                                 i_Safety_OK                := #io_System_Control.Safety_OK,
	                                 i_CMD_Reset                := #io_System_Control.OS_Reset,
	                                 i_CMD_Maintenance_Mode     := #io_Command.Man_Mode_Servo,
	                                 i_CMD_Disable_Axis         := #io_Command.Servo_Array[9].Man_Disable_Axis,
	                                 i_CMD_Home                 := #io_Command.Servo_Array[9].Man_Home,
	                                 i_CMD_Jog_Left             := #io_Command.Servo_Array[9].Man_Jog_Left,
	                                 i_CMD_Jog_Right            := #io_Command.Servo_Array[9].Man_Jog_Right,
	                                 i_CMD_Save                 := #io_Command.Servo_Array[9].Man_Save_Parameter,
	                                 i_CMD_Straight             := #s_Servo_Array_Command[9].CMD_Straight,
	                                 i_CMD_Divert_Left          := #s_Servo_Array_Command[9].CMD_Left,
	                                 i_CMD_Divert_Right         := #s_Servo_Array_Command[9].CMD_Right,
	                                 i_HW_Setting               := #i_Setting.Hardware.Servo_U481,
	                                 o_Ready_To_Reset           => #s_Servo_Ready_To_Reset[9],
	                                 o_ER_PN_Not_Present        => #s_Servo_Status[9].ER_PN_NotPresent,
	                                 o_ER_PN_Error              => #s_Servo_Status[9].ER_PN_Error,
	                                 o_ST_Axis_Enabled          => #s_Servo_Status[9].ST_Axis_Enabled,
	                                 o_ST_Position_Reached      => #s_Servo_Status[9].ST_Axis_Position_Reached,
	                                 o_OL_Maintenance_Mode      => #s_Servo_Status[9].OL_Maintenance_Mode,
	                                 o_ER_STO_Active            => #s_Servo_Status[9].ER_STO_Active,
	                                 o_WN_Motor_Alarm           => #s_Servo_Status[9].WN_Servo_Warn,
	                                 o_ER_Motor_Fault           => #s_Servo_Status[9].ER_Servo_Fault,
	                                 o_ER_Home_Position_Missing => #s_Servo_Status[9].ER_Home_Position_Missed,
	                                 o_ST_Act_Position          => #s_Servo_Status[9].ST_Act_Position,
	                                 o_AlarmCode                 => #s_Servo_Status[9].AlarmCode,
	                                 o_FaultCode                => #s_Servo_Status[9].ErrorCode,
	                                 io_Global                  := #io_Global,
	                                 io_S210_Interface          := #io_Interface.Servo9);
	    END_REGION
	END_REGION

	REGION NETWORK: Combine System Feedback Status
	    #io_System_Control.Ready_To_Reset := #s_Servo_Ready_To_Reset[1]
	    OR #s_Servo_Ready_To_Reset[2]
	    OR #s_Servo_Ready_To_Reset[3]
	    OR #s_Servo_Ready_To_Reset[4]
	    OR #s_Servo_Ready_To_Reset[5]
	    OR #s_Servo_Ready_To_Reset[6]
	    OR #s_Servo_Ready_To_Reset[7]
	    OR #s_Servo_Ready_To_Reset[8]
	    OR #s_Servo_Ready_To_Reset[9];
	END_REGION

	REGION Status Output

	    #o_Status.Roller_Module_1 := #s_Roller_Module_Status[1];
	    #o_Status.Roller_Module_2 := #s_Roller_Module_Status[2];
	    #o_Status.Roller_Module_3 := #s_Roller_Module_Status[3];
	    #o_Status.Roller_Module_4 := #s_Roller_Module_Status[4];
	    #o_Status.Roller_Module_5 := #s_Roller_Module_Status[5];
	    #o_Status.Roller_Module_6 := #s_Roller_Module_Status[6];
	    #o_Status.Roller_Module_7 := #s_Roller_Module_Status[7];
	    #o_Status.Roller_Module_8 := #s_Roller_Module_Status[8];
	    #o_Status.Roller_Module_9 := #s_Roller_Module_Status[9];

	    #o_Status.Servo_1 := #s_Servo_Status[1];
	    #o_Status.Servo_2 := #s_Servo_Status[2];
	    #o_Status.Servo_3 := #s_Servo_Status[3];
	    #o_Status.Servo_4 := #s_Servo_Status[4];
	    #o_Status.Servo_5 := #s_Servo_Status[5];
	    #o_Status.Servo_6 := #s_Servo_Status[6];
	    #o_Status.Servo_7 := #s_Servo_Status[7];
	    #o_Status.Servo_8 := #s_Servo_Status[8];
	    #o_Status.Servo_9 := #s_Servo_Status[9];

	    #o_General_Status.Safety_Stop := NOT #io_System_Control.Safety_OK;
	    #o_General_Status.Off_Line := #io_Command.Man_Mode_Servo OR #io_Command.Man_Mode;
	    #o_General_Status.Manual := #io_Command.Manual_Mode;
	    #o_General_Status.Error := #o_Status.ER_Modbus_Gateway_Initialize_Fault
	    OR #o_Status.ER_Modbus_Gateway_Communication_Fault
	    OR #s_Servo_Status[1].ER_PN_NotPresent
	    OR #s_Servo_Status[2].ER_PN_NotPresent
	    OR #s_Servo_Status[3].ER_PN_NotPresent
	    OR #s_Servo_Status[4].ER_PN_NotPresent
	    OR #s_Servo_Status[5].ER_PN_NotPresent
	    OR #s_Servo_Status[6].ER_PN_NotPresent
	    OR #s_Servo_Status[7].ER_PN_NotPresent
	    OR #s_Servo_Status[8].ER_PN_NotPresent
	    OR #s_Servo_Status[9].ER_PN_NotPresent
	    OR #s_Servo_Status[1].ER_Servo_Fault
	    OR #s_Servo_Status[2].ER_Servo_Fault
	    OR #s_Servo_Status[3].ER_Servo_Fault
	    OR #s_Servo_Status[4].ER_Servo_Fault
	    OR #s_Servo_Status[5].ER_Servo_Fault
	    OR #s_Servo_Status[6].ER_Servo_Fault
	    OR #s_Servo_Status[7].ER_Servo_Fault
	    OR #s_Servo_Status[8].ER_Servo_Fault
	    OR #s_Servo_Status[9].ER_Servo_Fault
	    OR #s_Servo_Status[1].ER_Home_Position_Missed
	    OR #s_Servo_Status[2].ER_Home_Position_Missed
	    OR #s_Servo_Status[3].ER_Home_Position_Missed
	    OR #s_Servo_Status[4].ER_Home_Position_Missed
	    OR #s_Servo_Status[5].ER_Home_Position_Missed
	    OR #s_Servo_Status[6].ER_Home_Position_Missed
	    OR #s_Servo_Status[7].ER_Home_Position_Missed
	    OR #s_Servo_Status[8].ER_Home_Position_Missed
	    OR #s_Servo_Status[9].ER_Home_Position_Missed
	    OR #s_Servo_Status[1].ER_STO_Active
	    OR #s_Servo_Status[2].ER_STO_Active
	    OR #s_Servo_Status[3].ER_STO_Active
	    OR #s_Servo_Status[4].ER_STO_Active
	    OR #s_Servo_Status[5].ER_STO_Active
	    OR #s_Servo_Status[6].ER_STO_Active
	    OR #s_Servo_Status[7].ER_STO_Active
	    OR #s_Servo_Status[8].ER_STO_Active
	    OR #s_Servo_Status[9].ER_STO_Active;

	    #o_General_Status.Warning := #s_Servo_Status[1].WN_Servo_Warn
	    OR #s_Servo_Status[2].WN_Servo_Warn
	    OR #s_Servo_Status[3].WN_Servo_Warn
	    OR #s_Servo_Status[4].WN_Servo_Warn
	    OR #s_Servo_Status[5].WN_Servo_Warn
	    OR #s_Servo_Status[6].WN_Servo_Warn
	    OR #s_Servo_Status[7].WN_Servo_Warn
	    OR #s_Servo_Status[8].WN_Servo_Warn
	    OR #s_Servo_Status[9].WN_Servo_Warn
	    OR #s_Roller_Module_Status[1].WN_Modbus_Com_Error
	    OR #s_Roller_Module_Status[1].WN_Motor_Blockage
	    OR #s_Roller_Module_Status[1].WN_Motor_NotConnected
	    OR #s_Roller_Module_Status[1].WN_Motor_NotHealthy
	    OR #s_Roller_Module_Status[2].WN_Modbus_Com_Error
	    OR #s_Roller_Module_Status[2].WN_Motor_Blockage
	    OR #s_Roller_Module_Status[2].WN_Motor_NotConnected
	    OR #s_Roller_Module_Status[2].WN_Motor_NotHealthy
	    OR #s_Roller_Module_Status[3].WN_Modbus_Com_Error
	    OR #s_Roller_Module_Status[3].WN_Motor_Blockage
	    OR #s_Roller_Module_Status[3].WN_Motor_NotConnected
	    OR #s_Roller_Module_Status[3].WN_Motor_NotHealthy
	    OR #s_Roller_Module_Status[4].WN_Modbus_Com_Error
	    OR #s_Roller_Module_Status[4].WN_Motor_Blockage
	    OR #s_Roller_Module_Status[4].WN_Motor_NotConnected
	    OR #s_Roller_Module_Status[4].WN_Motor_NotHealthy
	    OR #s_Roller_Module_Status[5].WN_Modbus_Com_Error
	    OR #s_Roller_Module_Status[5].WN_Motor_Blockage
	    OR #s_Roller_Module_Status[5].WN_Motor_NotConnected
	    OR #s_Roller_Module_Status[5].WN_Motor_NotHealthy
	    OR #s_Roller_Module_Status[6].WN_Modbus_Com_Error
	    OR #s_Roller_Module_Status[6].WN_Motor_Blockage
	    OR #s_Roller_Module_Status[6].WN_Motor_NotConnected
	    OR #s_Roller_Module_Status[6].WN_Motor_NotHealthy
	    OR #s_Roller_Module_Status[7].WN_Modbus_Com_Error
	    OR #s_Roller_Module_Status[7].WN_Motor_Blockage
	    OR #s_Roller_Module_Status[7].WN_Motor_NotConnected
	    OR #s_Roller_Module_Status[7].WN_Motor_NotHealthy
	    OR #s_Roller_Module_Status[8].WN_Modbus_Com_Error
	    OR #s_Roller_Module_Status[8].WN_Motor_Blockage
	    OR #s_Roller_Module_Status[8].WN_Motor_NotConnected
	    OR #s_Roller_Module_Status[8].WN_Motor_NotHealthy
	    OR #s_Roller_Module_Status[9].WN_Modbus_Com_Error
	    OR #s_Roller_Module_Status[9].WN_Motor_Blockage
	    OR #s_Roller_Module_Status[9].WN_Motor_NotConnected
	    OR #s_Roller_Module_Status[9].WN_Motor_NotHealthy;
	END_REGION

END_FUNCTION_BLOCK

TYPE "UDT_ADTA_Interface"
VERSION : 0.1
   STRUCT
      Input : Struct
         Spare_0_0 : Bool;
         Spare_0_1 : Bool;
         Spare_0_2 : Bool;
         Spare_0_3 : Bool;
         Spare_0_4 : Bool;
         Spare_0_5 : Bool;
         Spare_0_6 : Bool;
         Spare_0_7 : Bool;
         Spare_1_0 : Bool;
         Spare_1_1 : Bool;
         Spare_1_2 : Bool;
         Spare_1_3 : Bool;
         Spare_1_4 : Bool;
         Spare_1_5 : Bool;
         Spare_1_6 : Bool;
         Spare_1_7 : Bool;
         Spare_Byte_2 : Byte;
         Spare_Byte_3 : Byte;
         Spare_Byte_4 : Byte;
         Spare_Byte_5 : Byte;
         Spare_Byte_6 : Byte;
         Spare_Byte_7 : Byte;
         Spare_Byte_8 : Byte;
         Spare_Byte_9 : Byte;
         Spare_Byte_10 : Byte;
         Spare_Byte_11 : Byte;
         Spare_Byte_12 : Byte;
         Spare_Byte_13 : Byte;
         Spare_Byte_14 : Byte;
         Spare_Byte_15 : Byte;
      END_STRUCT;
      Output : Struct
         Spare_0_0 : Bool;
         Spare_0_1 : Bool;
         Spare_0_2 : Bool;
         Spare_0_3 : Bool;
         Spare_0_4 : Bool;
         Spare_0_5 : Bool;
         Spare_0_6 : Bool;
         Spare_0_7 : Bool;
         Spare_1_0 : Bool;
         Spare_1_1 : Bool;
         Spare_1_2 : Bool;
         Spare_1_3 : Bool;
         Spare_1_4 : Bool;
         Spare_1_5 : Bool;
         Spare_1_6 : Bool;
         Spare_1_7 : Bool;
         Spare_Byte_2 : Byte;
         Spare_Byte_3 : Byte;
         Spare_Byte_4 : Byte;
         Spare_Byte_5 : Byte;
         Spare_Byte_6 : Byte;
         Spare_Byte_7 : Byte;
         Spare_Byte_8 : Byte;
         Spare_Byte_9 : Byte;
         Spare_Byte_10 : Byte;
         Spare_Byte_11 : Byte;
         Spare_Byte_12 : Byte;
         Spare_Byte_13 : Byte;
         Spare_Byte_14 : Byte;
         Spare_Byte_15 : Byte;
      END_STRUCT;
   END_STRUCT;

END_TYPE

TYPE "UDT_Jam_Addon_IO"
VERSION : 0.1
   STRUCT
      Reset_Btn : Bool;
      Jam_Active : Bool;
   END_STRUCT;

END_TYPE

TYPE "UDT_NBS_Interface"
VERSION : 0.1
   STRUCT
      Input : Struct
         CMD_Start : Bool;
         CMD_Stop : Bool;
         CMD_Reset : Bool;
         Infeed_RTR : Bool;
         Speed1 : Bool;
         PassThrough_Mode : Bool;
         EngergySaving : Bool;
         Outfeed_RTS : Bool;
         LifeSign : Bool;
         Speed2 : Bool;
         Gap1 : Bool;
         Gap2 : Bool;
         Gap3 : Bool;
         Spare_1_5 : Bool;
         Spare_1_6 : Bool;
         Spare_1_7 : Bool;
         Spare_Byte_2 : Byte;
         Spare_Byte_3 : Byte;
         Spare_Byte_4 : Byte;
         Spare_Byte_5 : Byte;
         Spare_Byte_6 : Byte;
         Spare_Byte_7 : Byte;
         Spare_Byte_8 : Byte;
         Spare_Byte_9 : Byte;
         Spare_Byte_10 : Byte;
         Spare_Byte_11 : Byte;
         Spare_Byte_12 : Byte;
         Spare_Byte_13 : Byte;
         Spare_Byte_14 : Byte;
         Spare_Byte_15 : Byte;
      END_STRUCT;
      Output : Struct
         Infeed_RTS : Bool;
         Chute_RTR : Bool;
         LifeSign : Bool;
         Spare_0_3 : Bool;
         Spare_0_4 : Bool;
         Spare_0_5 : Bool;
         Spare_0_6 : Bool;
         Spare_0_7 : Bool;
         Spare_1_0 : Bool;
         Spare_1_1 : Bool;
         Spare_1_2 : Bool;
         Spare_1_3 : Bool;
         Spare_1_4 : Bool;
         Spare_1_5 : Bool;
         Spare_1_6 : Bool;
         Spare_1_7 : Bool;
         Spare_Byte_2 : Byte;
         Spare_Byte_3 : Byte;
         Spare_Byte_4 : Byte;
         Spare_Byte_5 : Byte;
         Spare_Byte_6 : Byte;
         Spare_Byte_7 : Byte;
         Spare_Byte_8 : Byte;
         Spare_Byte_9 : Byte;
         Spare_Byte_10 : Byte;
         Spare_Byte_11 : Byte;
         Spare_Byte_12 : Byte;
         Spare_Byte_13 : Byte;
         Spare_Byte_14 : Byte;
         Spare_Byte_15 : Byte;
      END_STRUCT;
   END_STRUCT;

END_TYPE

TYPE "UDT_Merge_Singulator_Interface"
VERSION : 0.1
   STRUCT
      Input : Struct
         OperateMode : Bool;   // False: singulate mode True: passthrough mode
         LowCapacityMode : Bool;   // False: high capacity singulate mode True: low capacity singulate mode
         ManualMode : Bool;   // False: auto mode True: manual mode
         RunningState : Bool;   // False: stopped True: running
         DeviceNoFault : Bool;   // False: fault True: ok
         DeviceNoEmergencyStop : Bool;   // False: emerengency stop True: ok
         LeftInfeed_RTR : Bool;   // Left infeed ready to receive
         RightInfeed_RTR : Bool;   // Right infeed ready to receive
         OutfeedRTS : Bool;
         NoJam : Bool;   // False: jam True: ok
         SingulateWarn : Bool;   // Singulate ratio < 97%
         SingulateFault : Bool;   // Singulate ratio < 95%
         Spare_1_4 : Bool;
         Spare_1_5 : Bool;
         Spare_1_6 : Bool;
         Spare_1_7 : Bool;
         Spare_Byte_2 : Byte;
         Spare_Byte_3 : Byte;
         Spare_Byte_4 : Byte;
         Spare_Byte_5 : Byte;
         Spare_Byte_6 : Byte;
         Spare_Byte_7 : Byte;
         Spare_Byte_8 : Byte;
         Spare_Byte_9 : Byte;
         Spare_Byte_10 : Byte;
         Spare_Byte_11 : Byte;
         Spare_Byte_12 : Byte;
         Spare_Byte_13 : Byte;
         Spare_Byte_14 : Byte;
         Spare_Byte_15 : Byte;
      END_STRUCT;
      Output : Struct
         Enable : Bool;
         ActivatePassthroughMode : Bool;
         ActivateLowCapacityMode : Bool;
         OutfeedRTR : Bool;
         NoEmergencyStop : Bool;
         Reset : Bool;
         LeftInfeed_PE : Bool;
         RightInfeed_PE : Bool;
         Speed1 : Bool;
         Speed2 : Bool;
         Gap1 : Bool;
         Gap2 : Bool;
         Gap3 : Bool;
         Outfeed_PE : Bool;
         LeftInfeed_RTS : Bool;
         RightInfeed_RTS : Bool;
         Spare_Byte_2 : Byte;
         Spare_Byte_3 : Byte;
         Spare_Byte_4 : Byte;
         Spare_Byte_5 : Byte;
         Infeed_Left_Gen_Status : Word;
         Infeed_Right_Gen_Status : Word;
         Outfeed_Gen_Status : Word;
         Outfeed_Item_Len : Int;
         Outfeed_Items_Gap : Int;
      END_STRUCT;
   END_STRUCT;

END_TYPE

TYPE "UDT_Tipper_Interface"
VERSION : 0.1
   STRUCT
      Input : Struct
         Spare_0_0 : Bool;
         Spare_0_1 : Bool;
         Spare_0_2 : Bool;
         Spare_0_3 : Bool;
         Spare_0_4 : Bool;
         Spare_0_5 : Bool;
         Spare_0_6 : Bool;
         Spare_0_7 : Bool;
         Spare_1_0 : Bool;
         Spare_1_1 : Bool;
         Spare_1_2 : Bool;
         Spare_1_3 : Bool;
         Spare_1_4 : Bool;
         Spare_1_5 : Bool;
         Spare_1_6 : Bool;
         Spare_1_7 : Bool;
         Spare_Byte_2 : Byte;
         Spare_Byte_3 : Byte;
         Spare_Byte_4 : Byte;
         Spare_Byte_5 : Byte;
         Spare_Byte_6 : Byte;
         Spare_Byte_7 : Byte;
         Spare_Byte_8 : Byte;
         Spare_Byte_9 : Byte;
         Spare_Byte_10 : Byte;
         Spare_Byte_11 : Byte;
         Spare_Byte_12 : Byte;
         Spare_Byte_13 : Byte;
         Spare_Byte_14 : Byte;
         Spare_Byte_15 : Byte;
      END_STRUCT;
      Output : Struct
         Spare_0_0 : Bool;
         Spare_0_1 : Bool;
         Spare_0_2 : Bool;
         Spare_0_3 : Bool;
         Spare_0_4 : Bool;
         Spare_0_5 : Bool;
         Spare_0_6 : Bool;
         Spare_0_7 : Bool;
         Spare_1_0 : Bool;
         Spare_1_1 : Bool;
         Spare_1_2 : Bool;
         Spare_1_3 : Bool;
         Spare_1_4 : Bool;
         Spare_1_5 : Bool;
         Spare_1_6 : Bool;
         Spare_1_7 : Bool;
         Spare_Byte_2 : Byte;
         Spare_Byte_3 : Byte;
         Spare_Byte_4 : Byte;
         Spare_Byte_5 : Byte;
         Spare_Byte_6 : Byte;
         Spare_Byte_7 : Byte;
         Spare_Byte_8 : Byte;
         Spare_Byte_9 : Byte;
         Spare_Byte_10 : Byte;
         Spare_Byte_11 : Byte;
         Spare_Byte_12 : Byte;
         Spare_Byte_13 : Byte;
         Spare_Byte_14 : Byte;
         Spare_Byte_15 : Byte;
      END_STRUCT;
   END_STRUCT;

END_TYPE

TYPE "UDT_Echelon_Interface"
VERSION : 0.1
   STRUCT
      Input : Struct
         Ready_To_Receive : Bool;
         Ready_To_Send : Bool;
         Hold_Actuve : Bool;
         Slow_Mode_Active : Bool;
         Clearing_Active : Bool;
         Clearing_Completed : Bool;
         Spare_0_6 : Bool;   // Signal Spare Bit
         Spare_0_7 : Bool;   // Signal Spare Bit
         Spare_1_0 : Bool;   // Signal Spare Bit
         Spare_1_1 : Bool;   // Signal Spare Bit
         Spare_1_2 : Bool;   // Signal Spare Bit
         Spare_1_3 : Bool;   // Signal Spare Bit
         Spare_1_4 : Bool;   // Signal Spare Bit
         Spare_1_5 : Bool;   // Signal Spare Bit
         Spare_1_6 : Bool;   // Signal Spare Bit
         Spare_1_7 : Bool;   // Signal Spare Bit
         Spare_2_0 : Bool;   // Signal Spare Bit
         Spare_2_1 : Bool;   // Signal Spare Bit
         Spare_2_2 : Bool;   // Signal Spare Bit
         Spare_2_3 : Bool;   // Signal Spare Bit
         Spare_2_4 : Bool;   // Signal Spare Bit
         Spare_2_5 : Bool;   // Signal Spare Bit
         Spare_2_6 : Bool;   // Signal Spare Bit
         Spare_2_7 : Bool;   // Signal Spare Bit
         LifeSign : Bool;   // Heartbeat Signal (500ms)
         Spare_3_1 : Bool;   // Signal Spare Bit
         Spare_3_2 : Bool;   // Signal Spare Bit
         Spare_3_3 : Bool;   // Signal Spare Bit
         Spare_3_4 : Bool;   // Signal Spare Bit
         Spare_3_5 : Bool;   // Signal Spare Bit
         Spare_3_6 : Bool;   // Signal Spare Bit
         Spare_3_7 : Bool;   // Signal Spare Bit
         Running : Bool;
         Faulted : Bool;
         Spare_4_2 : Bool;   // Diagnostic Spare Bit
         Spare_4_3 : Bool;   // Diagnostic Spare Bit
         Spare_4_4 : Bool;   // Diagnostic Spare Bit
         Spare_4_5 : Bool;   // Diagnostic Spare Bit
         Energy_Saveing : Bool;
         Automatic_Mode : Bool;
         Manual_Mode : Bool;
         Maintenance_Mode : Bool;
         Jammed : Bool;
         Spare_5_3 : Bool;   // Diagnostic Spare Bit
         Spare_5_4 : Bool;   // Diagnostic Spare Bit
         Spare_5_5 : Bool;   // Diagnostic Spare Bit
         Spare_5_6 : Bool;   // Diagnostic Spare Bit
         Spare_5_7 : Bool;   // Diagnostic Spare Bit
         Spare_6_0 : Bool;   // Diagnostic Spare Bit
         Spare_6_1 : Bool;   // Diagnostic Spare Bit
         Spare_6_2 : Bool;   // Diagnostic Spare Bit
         Spare_6_3 : Bool;   // Diagnostic Spare Bit
         Spare_6_4 : Bool;   // Diagnostic Spare Bit
         Spare_6_5 : Bool;   // Diagnostic Spare Bit
         Spare_6_6 : Bool;   // Diagnostic Spare Bit
         Spare_6_7 : Bool;   // Diagnostic Spare Bit
         Spare_7_0 : Bool;   // Diagnostic Spare Bit
         Spare_7_1 : Bool;   // Diagnostic Spare Bit
         Spare_7_2 : Bool;   // Diagnostic Spare Bit
         Spare_7_3 : Bool;   // Diagnostic Spare Bit
         Spare_7_4 : Bool;   // Diagnostic Spare Bit
         Spare_7_5 : Bool;   // Diagnostic Spare Bit
         Spare_7_6 : Bool;   // Diagnostic Spare Bit
         Spare_7_7 : Bool;   // Diagnostic Spare Bit
         Infeed_Speed : Real;   // [m/s]
         Outfeed_Speed : Real;   // [m/s]
         Spare_16_0 : Real;   // RealValue Spare Data
         Spare_20_0 : Real;   // RealValue Spare Data
         Spare_24_0 : Real;   // RealValue Spare Data
         Spare_28_0 : Real;   // RealValue Spare Data
         Spare_32_0 : Real;   // RealValue Spare Data
         Spare_36_0 : Real;   // RealValue Spare Data
      END_STRUCT;
      Output : Struct
         Start_Command : Bool;
         Stop_Command : Bool;
         Reset_Alarm : Bool;
         Slow_Down : Bool;
         Wake_Up : Bool;
         Hold : Bool;
         Spare_0_6 : Bool;   // Signal Spare Bit
         Spare_0_7 : Bool;   // Signal Spare Bit
         Upstream_RTS : Bool;
         Downstream_RTR : Bool;
         Spare_1_2 : Bool;   // Signal Spare Bit
         Spare_1_3 : Bool;   // Signal Spare Bit
         Spare_1_4 : Bool;   // Signal Spare Bit
         Spare_1_5 : Bool;   // Signal Spare Bit
         Spare_1_6 : Bool;   // Signal Spare Bit
         Spare_1_7 : Bool;   // Signal Spare Bit
         Spare_2_0 : Bool := false;   // Signal Spare Bit
         Spare_2_1 : Bool := false;   // Signal Spare Bit
         Spare_2_2 : Bool := false;   // Signal Spare Bit
         Spare_2_3 : Bool := false;   // Signal Spare Bit
         Spare_2_4 : Bool := false;   // Signal Spare Bit
         Spare_2_5 : Bool := false;   // Signal Spare Bit
         Spare_2_6 : Bool := false;   // Signal Spare Bit
         Spare_2_7 : Bool := false;   // Signal Spare Bit
         LifeSign : Bool := false;   // Heartbeat Signal (500ms)
         Spare_3_1 : Bool := false;   // Signal Spare Bit
         Spare_3_2 : Bool := false;   // Signal Spare Bit
         Spare_3_3 : Bool := false;   // Signal Spare Bit
         Spare_3_4 : Bool := false;   // Signal Spare Bit
         Spare_3_5 : Bool := false;   // Signal Spare Bit
         Spare_3_6 : Bool := false;   // Signal Spare Bit
         Spare_3_7 : Bool := false;   // Signal Spare Bit
         Upstream_Running : Bool := false;
         Downstream_Running : Bool := false;
         Upstream_Faulted : Bool := false;
         Dowstream_Faulted : Bool := false;
         Spare_4_4 : Bool := false;   // Diagnostic Spare Bit
         Spare_4_5 : Bool := false;   // Diagnostic Spare Bit
         Spare_4_6 : Bool := false;   // Diagnostic Spare Bit
         Spare_4_7 : Bool := false;   // Diagnostic Spare Bit
         Spare_5_0 : Bool := false;   // Diagnostic Spare Bit
         Spare_5_1 : Bool := false;   // Diagnostic Spare Bit
         Spare_5_2 : Bool := false;   // Diagnostic Spare Bit
         Spare_5_3 : Bool := false;   // Diagnostic Spare Bit
         Spare_5_4 : Bool := false;   // Diagnostic Spare Bit
         Spare_5_5 : Bool := false;   // Diagnostic Spare Bit
         Spare_5_6 : Bool := false;   // Diagnostic Spare Bit
         Spare_5_7 : Bool := false;   // Diagnostic Spare Bit
         Spare_6_0 : Bool := false;   // Diagnostic Spare Bit
         Spare_6_1 : Bool := false;   // Diagnostic Spare Bit
         Spare_6_2 : Bool := false;   // Diagnostic Spare Bit
         Spare_6_3 : Bool := false;   // Diagnostic Spare Bit
         Spare_6_4 : Bool := false;   // Diagnostic Spare Bit
         Spare_6_5 : Bool := false;   // Diagnostic Spare Bit
         Spare_6_6 : Bool := false;   // Diagnostic Spare Bit
         Spare_6_7 : Bool := false;   // Diagnostic Spare Bit
         Spare_7_0 : Bool := false;   // Diagnostic Spare Bit
         Spare_7_1 : Bool := false;   // Diagnostic Spare Bit
         Spare_7_2 : Bool := false;   // Diagnostic Spare Bit
         Spare_7_3 : Bool := false;   // Diagnostic Spare Bit
         Spare_7_4 : Bool := false;   // Diagnostic Spare Bit
         Spare_7_5 : Bool := false;   // Diagnostic Spare Bit
         Spare_7_6 : Bool := false;   // Diagnostic Spare Bit
         Spare_7_7 : Bool := false;   // Diagnostic Spare Bit
         Infeed_Speed : Real := 0.0;   // [m/s]
         Outfeed_Speed : Real := 0.0;   // [m/s]
         Spare_16_0 : Real := 0.0;   // RealValue Spare Data
         Spare_20_0 : Real := 0.0;   // RealValue Spare Data
         Spare_24_0 : Real := 0.0;   // RealValue Spare Data
         Spare_28_0 : Real := 0.0;   // RealValue Spare Data
         Spare_32_0 : Real := 0.0;   // RealValue Spare Data
         Spare_36_0 : Real := 0.0;   // RealValue Spare Data
      END_STRUCT;
   END_STRUCT;

END_TYPE

TYPE "UDT_TL70_IO"
VERSION : 0.1
   STRUCT
      Module_1_Color : Int;   // 0 = Green, 1 = Red, 2 = Orange, 3 = Amber, 4 = Yellow, 5 = Lime Green, 6 = Spring Green, 7 = Cyan, 8 = Sky Blue, 9 = Blue, 10 = Violet, 11 = Magenta, 12 = Rose, 13 = Daylight White (5000K), 14 = Custom 1, 15 = Custom 2
      Module_1_Flash : Int;   // 0 = Off, 1 = Steady, 2 = Flash 1Hz, 3 = Flash 2Hz, 4 = Flash 10Hz, 5 = Flash Custom Rate
      Module_2_Color : Int;   // 0 = Green, 1 = Red, 2 = Orange, 3 = Amber, 4 = Yellow, 5 = Lime Green, 6 = Spring Green, 7 = Cyan, 8 = Sky Blue, 9 = Blue, 10 = Violet, 11 = Magenta, 12 = Rose, 13 = Daylight White (5000K), 14 = Custom 1, 15 = Custom 2
      Module_2_Flash : Int;   // 0 = Off, 1 = Steady, 2 = Flash 1Hz, 3 = Flash 2Hz, 4 = Flash 10Hz, 5 = Flash Custom Rate
      Module_3_Color : Int;   // 0 = Green, 1 = Red, 2 = Orange, 3 = Amber, 4 = Yellow, 5 = Lime Green, 6 = Spring Green, 7 = Cyan, 8 = Sky Blue, 9 = Blue, 10 = Violet, 11 = Magenta, 12 = Rose, 13 = Daylight White (5000K), 14 = Custom 1, 15 = Custom 2
      Module_3_Flash : Int;   // 0 = Off, 1 = Steady, 2 = Flash 1Hz, 3 = Flash 2Hz, 4 = Flash 10Hz, 5 = Flash Custom Rate
      Module_4_Color : Int;   // 0 = Green, 1 = Red, 2 = Orange, 3 = Amber, 4 = Yellow, 5 = Lime Green, 6 = Spring Green, 7 = Cyan, 8 = Sky Blue, 9 = Blue, 10 = Violet, 11 = Magenta, 12 = Rose, 13 = Daylight White (5000K), 14 = Custom 1, 15 = Custom 2
      Module_4_Flash : Int;   // 0 = Off, 1 = Steady, 2 = Flash 1Hz, 3 = Flash 2Hz, 4 = Flash 10Hz, 5 = Flash Custom Rate
      Module_5_Color : Int;   // 0 = Green, 1 = Red, 2 = Orange, 3 = Amber, 4 = Yellow, 5 = Lime Green, 6 = Spring Green, 7 = Cyan, 8 = Sky Blue, 9 = Blue, 10 = Violet, 11 = Magenta, 12 = Rose, 13 = Daylight White (5000K), 14 = Custom 1, 15 = Custom 2
      Module_5_Flash : Int;   // 0 = Off, 1 = Steady, 2 = Flash 1Hz, 3 = Flash 2Hz, 4 = Flash 10Hz, 5 = Flash Custom Rate
      Buzzer : Bool;
      Port_Healthy : Bool;
   END_STRUCT;

END_TYPE

TYPE "UDT_MCC_Command"
VERSION : 0.1
   STRUCT
      Start : Bool;
      Stop : Bool;
      Reset : Bool;
   END_STRUCT;

END_TYPE

TYPE "UDT_SCADA_Command"
VERSION : 0.1
   STRUCT
      Start : Bool;
      Stop : Bool;
      Reset : Bool;
   END_STRUCT;

END_TYPE

FUNCTION_BLOCK "FB_Conv_Dual_G115D"
{ S7_Optimized_Access := 'TRUE' }
VERSION : 0.1
   VAR_INPUT
      i_U01_Telegram_HW_ID : HW_SUBMODULE;
      i_U01_Additional_HW_ID : HW_SUBMODULE;
      i_U02_Telegram_HW_ID : HW_SUBMODULE;
      i_U02_Additional_HW_ID : HW_SUBMODULE;
      i_IO_PEC_Position : Bool;
      i_IO_PEC_Trigger : Bool;
      i_Setting : "UDT_Conv_Dual_G115D_Setting";
      i_External_Request : "UDT_External_Request";
      i_Command : "UDT_Conv_Dual_G115D_Command";
   END_VAR

   VAR_OUTPUT RETAIN
      o_Status : "UDT_Conv_Dual_G115D_Status";
      o_General_Status : "UDT_General_Status";
      o_Diagnostics : "UDT_Conv_Dual_G115D_Diagnostics";
   END_VAR

   VAR_IN_OUT
      io_Global : "UDT_Global";
      io_System_Control : "UDT_System_Control";
      io_U01_G115D_IO : "UDT_G115D_HW_Interface";
      io_U02_G115D_IO : "UDT_G115D_HW_Interface";
      io_FIF_Upstream : "UDT_Flow_Interface";
      io_FIF : "UDT_Flow_Interface";
      io_FIF_Downstream : "UDT_Flow_Interface";
   END_VAR

   VAR
      s_FB_Displacement_AccDec : "FB_Displacement_AccDec";
      s_FB_EQP_PEC_Position : "FB_EQP_PEC_Position";
      s_FB_EQP_PEC_Trigger : "FB_EQP_PEC_Trigger";
      s_FB_EQP_Transport : "FB_EQP_Transport";
      s_U01_FB_HW_VFD_G115D : "FB_HW_VFD_G115D";
      s_U02_FB_HW_VFD_G115D : "FB_HW_VFD_G115D";
   END_VAR
   VAR RETAIN
      s_Cnt_PEC_Items : Int;
      s_Speed_Select : Int;
      s_SW_Actual_Speed : Int;
      s_U01_HW_Actual_Speed : Int;
      s_U02_HW_Actual_Speed : Int;
      s_CMD_PEC_Preset_Latch : Bool;
      s_CMD_Motor : Bool;
      s_CMD_Motor_Reverse : Bool;
      s_U01_HW_Req_Halt : Bool;
      s_U02_HW_Req_Halt : Bool;
      s_PE_Position_Latch : Bool;
      s_PE_Trigger_Latch : Bool;
      s_Ext_Req_Stop : Bool;
      s_Ext_Req_Halt : Bool;
      s_Ext_Req_Disable_Send : Bool;
      s_Ext_Req_Disable_Recv : Bool;
      s_Ext_Req_Rest_ESave : Bool;
      s_Ext_Req_Clear_Data : Bool;
      s_SW_Motor_OnSpeed : Bool;
      s_U01_HW_Motor_Running : Bool;
      s_U02_HW_Motor_Running : Bool;
   END_VAR

   VAR_TEMP
      t_PEC_Position_Items : UDInt;
      t_PEC_Trigger_Items : UDInt;
      t_PEC_Position_Ready_To_Reset : Bool;
      t_PEC_Trigger_Ready_To_Reset : Bool;
      t_U01_HW_VFD_Ready_To_Reset : Bool;
      t_U02_HW_VFD_Ready_To_Reset : Bool;
   END_VAR


BEGIN
	REGION NETWORK AA: Conveyor Cycle Displacement
	    #s_FB_Displacement_AccDec(i_Conveyor_Speed   := #io_FIF.Speed,
	                              i_Accelaration     := #i_Setting.Hardware_U01.Acceleration,
	                              i_Decelaration     := #i_Setting.Hardware_U01.Deceleration,
	                              i_Prev_Cycle_Time  := #io_Global.OB_Prev_Cycle_Time,
	                              i_PPI_Displacement := 0,
	                              i_Section_Run      := #io_FIF.Motor_Run,
	                              o_Motor_On_Speed   => #o_General_Status.Motor_On_Speed,
	                              o_Motor_Stopped    => #io_FIF.Motor_Stopped,
	                              o_Actual_Speed     => #s_SW_Actual_Speed,
	                              o_Displacement     => #io_FIF.Displacement);

	    #o_General_Status.Motor_Stopped := #io_FIF.Motor_Stopped;
	END_REGION

	REGION NETWORK BA: Equipment layer - PEC
	    #s_FB_EQP_PEC_Position(i_IO_Available             := #io_System_Control.IO_Available,
	                           i_CMD_Reset                := #io_System_Control.OS_Reset_Jam,
	                           i_CMD_Clear_Stat           := #io_System_Control.OS_Clear_Statistics,
	                           i_CFG_Blockage_Length      := #i_Setting.PE1.Blockage_Length,
	                           i_CFG_Delay_On             := #i_Setting.PE1.Delay_On,
	                           i_CFG_Delay_Off            := #i_Setting.PE1.Delay_Off,
	                           i_CFG_Shifting_Offset      := #i_Setting.PE1.Shifting_Offset,
	                           i_CFG_Handover_Offset      := #i_Setting.PE1.Handover_Offset,
	                           i_CFG_Detect_PEC_OnStopped := #i_Setting.PE1.Detect_PEC_OnStopped,
	                           i_CFG_Reset_Block_PEC_Oc   := #i_Setting.PE1.Reset_Block_PEC_Oc,
	                           i_CFG_Item_On              := #i_Setting.PE1.Item_On,
	                           i_CMD_Preset_Latch         := #s_CMD_PEC_Preset_Latch,
	                           i_CMD_Clear_Data           := #s_Ext_Req_Clear_Data,
	                           i_Cycle_Count              := #io_FIF.Displacement,
	                           i_IO_PEC                   := #i_IO_PEC_Position,
	                           i_Section_Running          := NOT #io_FIF.Motor_Stopped,
	                           o_Ready_To_Reset           => #t_PEC_Position_Ready_To_Reset,
	                           o_ER_PEC_Blockage          => #o_Status.ER_PE1_Blockage,
	                           o_PEC_Filter               => #s_PE_Position_Latch,
	                           o_Handover                 => #io_FIF.Handover,
	                           o_Cnt_Buffer_Used          => #s_Cnt_PEC_Items,
	                           o_Stat_Items               => #t_PEC_Position_Items);

	    #s_FB_EQP_PEC_Trigger(i_IO_Available             := #io_System_Control.IO_Available,
	                          i_CMD_Reset                := #io_System_Control.OS_Reset_Jam,
	                          i_CMD_Clear_Stat           := #io_System_Control.OS_Clear_Statistics,
	                          i_CFG_Blockage_Length      := #i_Setting.PE2.Blockage_Length,
	                          i_CFG_Delay_On             := #i_Setting.PE2.Delay_On,
	                          i_CFG_Delay_Off            := #i_Setting.PE2.Delay_Off,
	                          i_CFG_Detect_PEC_OnStopped := #i_Setting.PE2.Detect_PEC_OnStopped,
	                          i_CFG_Reset_Block_PEC_Oc   := #i_Setting.PE2.Reset_Block_PEC_Oc,
	                          i_CFG_Item_On              := #i_Setting.PE2.Item_On,
	                          i_CMD_Preset_Latch         := false,
	                          i_Cycle_Count              := #io_FIF.Displacement,
	                          i_IO_PEC                   := #i_IO_PEC_Trigger,
	                          i_Section_Running          := NOT #io_FIF.Motor_Stopped,
	                          o_Ready_To_Reset           => #t_PEC_Trigger_Ready_To_Reset,
	                          o_ER_PEC_Blockage          => #o_Status.ER_PE2_Blockage,
	                          o_PEC_Filter               => #s_PE_Trigger_Latch,
	                          o_Stat_Items               => #t_PEC_Trigger_Items);

	    #io_FIF.PECTrigger_Latch := #s_PE_Trigger_Latch;
	END_REGION

	REGION NETWORK CA: Conditions to basic control
	    // Condition to request stop
	    #s_Ext_Req_Stop := #o_Status.ER_U01_VFD_PN_NotPresent
	    // OR #o_Status.ER_U01_PN_Error
	    OR #o_Status.ER_U01_VFD_Fault
	    OR #o_Status.ER_U01_VFD_STO_Active
	    OR #o_Status.ER_U02_VFD_PN_NotPresent
	    // OR #o_Status.ER_U02_PN_Error
	    OR #o_Status.ER_U02_VFD_Fault
	    OR #o_Status.ER_U02_VFD_STO_Active
	    OR #i_External_Request.Request_Stop;

	    // Condition to request halt
	    #s_Ext_Req_Halt := #s_U01_HW_Req_Halt
	    OR #s_U02_HW_Req_Halt
	    OR #i_External_Request.Request_Halt
	    OR #i_Command.Man_Mode
	    OR #o_Status.ER_PE1_Blockage
	    OR #o_Status.ER_PE2_Blockage;

	    // Condition to request disable send
	    #s_Ext_Req_Disable_Send := #i_External_Request.Request_Disable_Send;

	    // Condition to request disable receive
	    #s_Ext_Req_Disable_Recv := #i_External_Request.Request_Disable_Receive OR #i_Command.Man_Mode;

	    // Condition to request reset engergy saving
	    #s_Ext_Req_Rest_ESave := #i_External_Request.Request_Reset_EnergySave OR #io_Global.Common_Setting.Disable_Energy_Saving OR #i_Command.Cmd_Reset_ESave OR #s_PE_Trigger_Latch OR #s_FB_EQP_PEC_Position.s_PEC_Filter;

	    // Condition to request clear flow interface data
	    #s_Ext_Req_Clear_Data := #i_External_Request.Request_Clear_Data OR (#i_Command.Man_Clear AND #i_Command.Man_Mode);
	END_REGION

	REGION NETWORK DA: Equipment Layer - Basic
	    #s_FB_EQP_Transport(i_Enable                 := #io_System_Control.Enable,
	                        i_IO_Available           := #io_System_Control.IO_Available,
	                        i_Safety_OK              := #io_System_Control.Safety_OK,
	                        i_CMD_Reset              := #io_System_Control.OS_Reset,
	                        i_CMD_Start              := #io_System_Control.OS_Start,
	                        i_CMD_Controlled_Stop    := #io_System_Control.Controlled_Stop,
	                        i_End_PEC_Latch          := #s_PE_Position_Latch,
	                        i_Manual_Run             := #i_Command.Man_Run AND #i_Command.Man_Mode,
	                        i_CFG_Slave_Conveyor     := #i_Setting.Base_Conveyor.Slave_Mode,
	                        i_CFG_Enable_DieForward  := #i_Setting.Base_Conveyor.Enable_DieForward,
	                        i_Delay_Waiting_Item     := #i_Setting.Base_Conveyor.Delay_Waiting_Item,
	                        i_Delay_Dieback          := #i_Setting.Base_Conveyor.Delay_Dieback,
	                        i_Delay_Startup          := #i_Setting.Base_Conveyor.Delay_Startup,
	                        i_Delay_Finish_Handover  := #i_Setting.Base_Conveyor.Delay_Finish_Handover,
	                        i_Delay_Energysave       := #i_Setting.Base_Conveyor.Delay_Energysave,
	                        i_Delay_Cascade_Startup  := #i_Setting.Base_Conveyor.Delay_Cascade_Startup,
	                        i_Delay_Cascade_Shutdown := #i_Setting.Base_Conveyor.Delay_Cascade_Shutdown,
	                        i_Delay_Motor_Startup    := #i_Setting.Hardware_U01.Magnetization_Delay,
	                        i_Minimum_Gap            := #i_Setting.Flow_Control.Minimum_Gap,
	                        i_Minimum_Head_To_Head   := #i_Setting.Flow_Control.Minimum_Head_To_Head,
	                        i_Ext_Req_Stop           := #s_Ext_Req_Stop,
	                        i_Ext_Req_Halt           := #s_Ext_Req_Halt,
	                        i_Ext_Req_Dis_Send       := #s_Ext_Req_Disable_Send,
	                        i_Ext_Req_Dis_Recv       := #s_Ext_Req_Disable_Recv,
	                        i_Ext_Req_Rst_ESave      := #s_Ext_Req_Rest_ESave,
	                        i_Ext_Req_Clear_Data     := #s_Ext_Req_Clear_Data,
	                        o_Ready_To_Start         => #io_System_Control.Ready_To_Start,
	                        o_ST_Safety_Stop         => #o_General_Status.Safety_Stop,
	                        o_ST_Items               => #o_General_Status.Items,
	                        o_ST_Die_Back            => #o_General_Status.Die_Back,
	                        o_ST_Motor_Running       => #o_General_Status.Motor_Running,
	                        o_ST_Started             => #o_General_Status.Started,
	                        o_ST_Energy_Saving       => #o_General_Status.Energy_Saving,
	                        o_MTR_Run                => #s_CMD_Motor,
	                        io_Global                := #io_Global,
	                        io_FIF_Upstream          := #io_FIF_Upstream,
	                        io_FIF                   := #io_FIF,
	                        io_FIF_Downstream        := #io_FIF_Downstream);
	END_REGION

	REGION NETWORK EA: Hardware Layer - G115D Convertor
	    #s_Speed_Select := #i_External_Request.Request_Speed;

	    #s_U01_FB_HW_VFD_G115D(i_Telegram_HW_ID        := #i_U01_Telegram_HW_ID,
	                           i_Additional_HW_ID      := #i_U01_Additional_HW_ID,
	                           i_Enable                := (#io_System_Control.Enable OR #i_Command.Man_Mode) AND NOT #i_Command.Man_DisableAxis,
	                           i_IO_Available          := #io_System_Control.IO_Available,
	                           i_Safety_OK             := #io_System_Control.Safety_OK,
	                           i_CMD_Reset             := #io_System_Control.OS_Reset,
	                           i_CMD_Clear_Stat        := #io_System_Control.OS_Clear_Statistics,
	                           i_HW_Setting            := #i_Setting.Hardware_U01,
	                           i_CFG_Motor_Switch_Time := 500,
	                           i_CMD_Select_Speed      := #s_Speed_Select,
	                           i_CMD_Motor_Run         := #s_CMD_Motor,
	                           i_CMD_Motor_Reverse     := #s_CMD_Motor_Reverse,
	                           o_Ready_To_Reset        => #t_U01_HW_VFD_Ready_To_Reset,
	                           o_Req_Halt              => #s_U01_HW_Req_Halt,
	                           o_ER_PN_Not_Present     => #o_Status.ER_U01_VFD_PN_NotPresent,
	                           o_ER_PN_Error           => #o_Status.ER_U01_VFD_PN_Error,
	                           o_ER_Motor_Fault        => #o_Status.ER_U01_VFD_Fault,
	                           o_WN_Motor_Alarm        => #o_Status.WN_U01_VFD_Alarm,
	                           o_ER_STO_Active         => #o_Status.ER_U01_VFD_STO_Active,
	                           o_WN_No_MemoryCard      => #o_Status.WN_U01_No_MemoryCard,
	                           o_ST_Motor_Running      => #s_U01_HW_Motor_Running,
	                           o_FaultCode             => #o_Status.U01_FaultCode,
	                           o_AlarmCode             => #o_Status.U01_AlarmCode,
	                           o_Speed_Selected        => #io_FIF.Speed,
	                           o_Diagnostics           => #o_Diagnostics.Hardware_U01,
	                           io_Global               := #io_Global,
	                           io_G115D_Interface      := #io_U01_G115D_IO);
	END_REGION

	REGION NETWORK EB: Hardware Layer - G115D Convertor
	    #s_Speed_Select := #i_External_Request.Request_Speed;

	    #s_U02_FB_HW_VFD_G115D(i_Telegram_HW_ID        := #i_U02_Telegram_HW_ID,
	                           i_Additional_HW_ID      := #i_U02_Additional_HW_ID,
	                           i_Enable                := (#io_System_Control.Enable OR #i_Command.Man_Mode) AND NOT #i_Command.Man_DisableAxis,
	                           i_IO_Available          := #io_System_Control.IO_Available,
	                           i_Safety_OK             := #io_System_Control.Safety_OK,
	                           i_CMD_Reset             := #io_System_Control.OS_Reset,
	                           i_CMD_Clear_Stat        := #io_System_Control.OS_Clear_Statistics,
	                           i_HW_Setting            := #i_Setting.Hardware_U02,
	                           i_CFG_Motor_Switch_Time := 500,
	                           i_CMD_Select_Speed      := #s_Speed_Select,
	                           i_CMD_Motor_Run         := #s_CMD_Motor,
	                           i_CMD_Motor_Reverse     := #s_CMD_Motor_Reverse,
	                           o_Ready_To_Reset        => #t_U02_HW_VFD_Ready_To_Reset,
	                           o_Req_Halt              => #s_U02_HW_Req_Halt,
	                           o_ER_PN_Not_Present     => #o_Status.ER_U02_VFD_PN_NotPresent,
	                           o_ER_PN_Error           => #o_Status.ER_U02_VFD_PN_Error,
	                           o_ER_Motor_Fault        => #o_Status.ER_U02_VFD_Fault,
	                           o_WN_Motor_Alarm        => #o_Status.WN_U02_VFD_Alarm,
	                           o_ER_STO_Active         => #o_Status.ER_U02_VFD_STO_Active,
	                           o_WN_No_MemoryCard      => #o_Status.WN_U02_No_MemoryCard,
	                           o_ST_Motor_Running      => #s_U02_HW_Motor_Running,
	                           o_FaultCode             => #o_Status.U02_FaultCode,
	                           o_AlarmCode             => #o_Status.U02_AlarmCode,
	                           o_Diagnostics           => #o_Diagnostics.Hardware_U02,
	                           io_Global               := #io_Global,
	                           io_G115D_Interface      := #io_U02_G115D_IO);
	END_REGION

	REGION NETWORK: Diagnositcs
	    #o_Diagnostics.RTS := #io_FIF.RTS;
	    #o_Diagnostics.TIP := #io_FIF.TIP;
	    #o_Diagnostics.Downstream_RTR := #io_FIF_Downstream.RTR;
	    #o_Diagnostics.Displacement := #io_FIF.Displacement;
	    #o_Diagnostics.Items_Count := MAX_UDINT(IN1 := #t_PEC_Position_Items, IN2 := #t_PEC_Trigger_Items);
	END_REGION

	REGION NETWORK FA: Make Generate Status
	    #o_Status.OL_Maintenance_Mode := #i_Command.Man_Mode;

	    #o_General_Status.Safety_Stop := #o_Status.ER_U01_VFD_STO_Active OR #o_Status.ER_U02_VFD_STO_Active OR NOT #io_System_Control.Safety_OK;
	    #o_General_Status.Off_Line := #o_Status.OL_Maintenance_Mode;
	    #o_General_Status.Manual := FALSE;
	    #o_General_Status.Error := #o_Status.ER_U01_VFD_PN_NotPresent
	    OR #o_Status.ER_U01_VFD_PN_Error
	    OR #o_Status.ER_U01_VFD_Fault
	    OR #o_Status.ER_U02_VFD_PN_NotPresent
	    OR #o_Status.ER_U02_VFD_PN_Error
	    OR #o_Status.ER_U02_VFD_Fault;
	    #o_General_Status.Jam := #o_Status.ER_PE1_Blockage OR #o_Status.ER_PE2_Blockage;
	    #o_General_Status.Warning := #o_Status.WN_U01_VFD_Alarm
	    OR #o_Status.WN_U01_No_MemoryCard
	    OR #o_Status.WN_U02_VFD_Alarm
	    OR #o_Status.WN_U02_No_MemoryCard;
	END_REGION

	REGION NETWORK EA: System Feedback State
	    #io_System_Control.Ready_To_Reset := #t_PEC_Position_Ready_To_Reset
	    OR #t_PEC_Trigger_Ready_To_Reset
	    OR #t_U01_HW_VFD_Ready_To_Reset
	    OR #t_U02_HW_VFD_Ready_To_Reset;
	END_REGION
END_FUNCTION_BLOCK

TYPE "UDT_Chute_Status"
VERSION : 0.1
   STRUCT
      ER_Chute_Full : Bool;
      Spare_0_1 : Bool;
      Spare_0_2 : Bool;
      Spare_0_3 : Bool;
      Spare_0_4 : Bool;
      Spare_0_5 : Bool;
      Spare_0_6 : Bool;
      Spare_0_7 : Bool;
      Spare_1_0 : Bool;
      Spare_1_1 : Bool;
      Spare_1_2 : Bool;
      Spare_1_3 : Bool;
      Spare_1_4 : Bool;
      Spare_1_5 : Bool;
      Spare_1_6 : Bool;
      Spare_1_7 : Bool;
   END_STRUCT;

END_TYPE

